(* IEC 61131-3 sources: TetherPLC/tests/compat (part 2) *)

(* ---- tc2_mc2_case.st ---- *)
PROGRAM Tc2Mc2Case
VAR
    mask   AT %QD0 : DINT;
    st     : INT;
    ax     : FB_MotionAxis;
    axH    : UDINT;
    pwr    : MC_Power;
    rst    : MC_Reset;
    sp     : MC_SetPosition;
    rpos   : MC_ReadActualPosition;
    rvel   : MC_ReadActualVelocity;
    rerr   : MC_ReadAxisError;
    rstat  : MC_ReadStatus;
    enSig  : BOOL;
    rstExec: BOOL;
    spExec : BOOL;
    spPos  : DINT;
    spMode : BOOL;
END_VAR

// Create the simulated axis once (raw FB_MotionAxis OP=1).
IF st = 0 THEN
    ax.UNITS_PER_REV := 1000;
    ax.MAX_VEL := 1000;
    ax.MAX_ACCEL := 5000;
    ax.MAX_DECEL := 5000;
    ax.POS_MIN := -100000;
    ax.POS_MAX := 100000;
    ax.HOME_OFFSET := 0;
    ax.FOLLOW_WINDOW := 3;
    ax.FLAGS := 1;
    ax.OP := 1;
    ax();
    IF ax.AXIS <> 0 AND ax.STATUS = 0 THEN
        axH := ax.AXIS;
        mask := mask + 1;
    END_IF;
    st := 1;
END_IF;

// Command/select signals derived from st (each command state is a
// single scan, giving each Execute FB exactly one rising edge).
enSig   := (st >= 1) AND (st <= 7);   // powered through the reset
rstExec := (st = 6);
spExec  := (st = 2) OR (st = 4);
spPos   := 1000;
IF st = 4 THEN spPos := 500; END_IF;
spMode  := (st = 4);

// Drive every MC wrapper each scan.
pwr(Enable := enSig, Enable_Positive := TRUE,
    Enable_Negative := TRUE, Axis := axH);
rst(Execute := rstExec, Axis := axH);
sp(Execute := spExec, Position := spPos, Mode := spMode, Axis := axH);
rpos(Enable := TRUE, Axis := axH);
rvel(Enable := TRUE, Axis := axH);
rerr(Enable := TRUE, Axis := axH);
rstat(Enable := TRUE, Axis := axH);

IF st = 1 THEN
    // MC_Power enable: wait for Status (OperationEnabled, ~2 scans)
    IF pwr.Status THEN
        mask := mask + 2;
        st := 2;
    END_IF;
ELSIF st = 2 THEN
    // absolute MC_SetPosition to 1000 fired this scan
    IF sp.Done THEN mask := mask + 4; END_IF;
    st := 3;
ELSIF st = 3 THEN
    // verify absolute position readback == 1000
    IF rpos.Valid AND rpos.Position = 1000 THEN
        mask := mask + 8;
    END_IF;
    st := 4;
ELSIF st = 4 THEN
    // relative MC_SetPosition +500 -> 1500 fired this scan
    IF sp.Done THEN mask := mask + 16; END_IF;
    st := 5;
ELSIF st = 5 THEN
    // verify relative readback == 1500 and the read FBs are valid
    IF rpos.Valid AND rpos.Position = 1500 THEN
        mask := mask + 32;
    END_IF;
    IF rvel.Valid AND rerr.Valid AND rstat.Valid THEN
        mask := mask + 64;
    END_IF;
    st := 6;
ELSIF st = 6 THEN
    // MC_Reset Execute edge -> Done (axis stays enabled)
    IF rst.Done THEN mask := mask + 128; END_IF;
    st := 7;
ELSIF st = 7 THEN
    // reset release scan; keep waiting for power to drop next
    st := 8;
ELSIF st = 8 THEN
    // enSig now FALSE: MC_Power disabled the axis; wait for
    // Status=FALSE and OperatingState=Disabled (0)
    IF NOT pwr.Status THEN
        mask := mask + 256;
        st := 9;
    END_IF;
ELSIF st = 9 THEN
    IF rstat.OperatingState = 0 THEN
        mask := mask + 512;
        st := 10;
    END_IF;
END_IF;

END_PROGRAM

(* ---- tc2_mc2_drive_case.st ---- *)
PROGRAM Tc2Mc2DriveCase
VAR
    mask   AT %QD0 : DINT;
    st     : INT;
    prevSt : INT;
    pulse  : BOOL;
    ax     : FB_MotionAxis;
    axM    : UDINT;
    axS    : UDINT;
    pwrM   : MC_Power;
    pwrS   : MC_Power;
    mvV    : MC_MoveVelocity;
    hlt    : MC_Halt;
    info   : FB_ReadDriveInfo;
    coeWr  : FB_CoEWrite;
    coeRd  : FB_CoERead;
    coeCmd : FB_CoEExecuteCommand;
    setOff : FB_SetPositionOffset;
    delOff : FB_DeletePositionOffset;
    brk    : FB_BrakeControl;
    rdPar  : FB_ReadDriveParameter;
    rdPar2 : FB_ReadDriveParameter;
    ax8kBrk : FB_CoEAX8000BrakeControl;
    ax8kTst : FB_CoEAX8000BrakeTest;
    ax8kPrk : FB_CoEAX8000ParkAxis;
    elBrk  : FB_CoEEL72xxBrakeControl;
    elSet  : FB_CoEEL72xxSetPositionOffset;
    saw    : MC_ReadFlyingSawCharacteristics;
    soeRd  : FB_SoERead;
    soeWrPw: FB_SoEWritePassword;
    soeCmd : FB_SoEExecuteCommand;
    soeCmd2: FB_SoEExecuteCommand;
    soeCmdSt: FB_SoEReadCommandState;
    soeRst : FB_SoEReset;
    ax5kV  : FB_SoEAX5000ReadActMainVoltage;
    ax5kFw : FB_SoEAX5000FirmwareUpdate;
    gv     : MC_GearInVelo;
    gp     : MC_GearInPos;
    rvelS  : MC_ReadActualVelocity;
    rposS  : MC_ReadActualPosition;
    rposM  : MC_ReadActualPosition;
    enSig  : BOOL;
    mvVEx  : BOOL;
    gvEx   : BOOL;
    gpEx   : BOOL;
    hltEx  : BOOL;
    cmdErrSeen : BOOL;
    cmdDoneSeen : BOOL;
    tog     : BOOL;
END_VAR

// Create two simulated axes (master slave0, slave slave1).
IF st = 0 THEN
    ax.UNITS_PER_REV := 1000;
    ax.MAX_VEL := 2000;
    ax.MAX_ACCEL := 8000;
    ax.MAX_DECEL := 8000;
    ax.POS_MIN := -200000;
    ax.POS_MAX := 200000;
    ax.HOME_OFFSET := 0;
    ax.FOLLOW_WINDOW := 3;
    ax.FLAGS := 1;
    ax.OP := 1; ax();
    IF ax.AXIS <> 0 THEN axM := ax.AXIS; END_IF;
    ax.OP := 1; ax();
    IF ax.AXIS <> 0 THEN axS := ax.AXIS; END_IF;
    IF axM <> 0 AND axS <> 0 THEN
        mask := mask + 1;                       // bit0: two axes
    END_IF;
    st := 1;
    prevSt := 0;
END_IF;

IF st <> prevSt THEN pulse := TRUE; ELSE pulse := FALSE; END_IF;
prevSt := st;
tog := NOT tog;   // re-pulse helper for the command-state polls

enSig  := (st >= 1) AND (st <= 29);
mvVEx  := pulse AND (st = 26);       // master velocity for gear tests
gvEx   := (st >= 27) AND (st <= 28); // velocity gear held
gpEx   := (st = 29);                 // position gear one scan
hltEx  := pulse AND (st = 30);

pwrM(Enable := enSig, Enable_Positive := TRUE, Enable_Negative := TRUE,
    Axis := axM);
pwrS(Enable := enSig, Enable_Positive := TRUE, Enable_Negative := TRUE,
    Axis := axS);
mvV(Execute := mvVEx, ContinuousUpdate := FALSE, Velocity := 400,
    Acceleration := 8000, Deceleration := 8000, Axis := axM);
hlt(Execute := hltEx, Deceleration := 8000, Axis := axM);
gv(Execute := gvEx, RatioNumerator := 2, RatioDenominator := 1,
   Acceleration := 8000, Deceleration := 8000, Master := axM, Slave := axS);
gp(Execute := gpEx, RatioNumerator := 1, RatioDenominator := 1,
   Acceleration := 8000, Deceleration := 8000, Master := axM, Slave := axS);
rvelS(Enable := TRUE, Axis := axS);
rposS(Enable := TRUE, Axis := axS);
rposM(Enable := TRUE, Axis := axM);

IF st = 1 THEN
    IF pwrM.Status AND pwrS.Status THEN
        mask := mask + 2;                       // bit1: powered
        st := 2;
    END_IF;
ELSIF st = 2 THEN
    info(Execute := pulse, Axis := axM);
    IF info.Valid AND info.State > 0 THEN
        mask := mask + 4;                       // bit2: drive info
        st := 3;
    END_IF;
ELSIF st = 3 THEN
    coeWr(Execute := pulse, Index := 16#2003, Value := 7, Axis := axM);
    IF coeWr.Done THEN
        mask := mask + 8;                       // bit3: CoE write
        st := 4;
    END_IF;
ELSIF st = 4 THEN
    coeRd(Execute := pulse, Index := 16#2003, Axis := axM);
    IF coeRd.Done AND coeRd.Value = 7 THEN
        mask := mask + 16;                      // bit4: CoE readback
        st := 5;
    END_IF;
ELSIF st = 5 THEN
    coeCmd(Execute := pulse, Command := 42, Axis := axM);
    IF coeCmd.Done THEN
        mask := mask + 32;                      // bit5: CoE command
        st := 6;
    END_IF;
ELSIF st = 6 THEN
    setOff(Execute := pulse, Position := 5000.0, Relative := FALSE,
           Feedback := 0, Memory := 0, Axis := axM);
    IF setOff.Done THEN
        mask := mask + 64;                      // bit6: pos offset
        st := 7;
    END_IF;
ELSIF st = 7 THEN
    rdPar(Execute := pulse, ParameterNumber := 16#2002, Mode := 0,
          Interval := 0, Axis := axM);
    IF rdPar.Valid AND rdPar.Value = 5000 THEN
        mask := mask + 128;                     // bit7: offset=5000
        st := 8;
    END_IF;
ELSIF st = 8 THEN
    delOff(Execute := pulse, Feedback := 0, Memory := 0, Axis := axM);
    IF delOff.Done THEN
        mask := mask + 256;                     // bit8: offset del
        st := 9;
    END_IF;
ELSIF st = 9 THEN
    brk(Execute := pulse, Mode := 3, Axis := axM);
    IF brk.Done THEN
        mask := mask + 512;                     // bit9: brake ctrl
        st := 10;
    END_IF;
ELSIF st = 10 THEN
    ax8kBrk(Execute := pulse, Mode := 1, Axis := axM);
    IF ax8kBrk.Done THEN
        mask := mask + 1024;                    // bit10: ax8k brake
        st := 11;
    END_IF;
ELSIF st = 11 THEN
    ax8kTst(Execute := pulse, Axis := axM);
    IF ax8kTst.Succeeded THEN
        mask := mask + 2048;                    // bit11: brake test
        st := 12;
    END_IF;
ELSIF st = 12 THEN
    ax8kPrk(Execute := pulse, Mode := 1, Axis := axM);
    IF ax8kPrk.Done THEN
        mask := mask + 4096;                    // bit12: ax8k park
        st := 13;
    END_IF;
ELSIF st = 13 THEN
    rdPar2(Execute := pulse, ParameterNumber := 16#2004, Mode := 0,
           Interval := 0, Axis := axM);
    IF rdPar2.Valid AND rdPar2.Value = 1 THEN
        mask := mask + 8192;                    // bit13: park=1
        st := 14;
    END_IF;
ELSIF st = 14 THEN
    elBrk(Execute := pulse, Mode := 2, Axis := axM);
    IF elBrk.Done THEN
        mask := mask + 16384;                   // bit14: el72xx brk
        st := 15;
    END_IF;
ELSIF st = 15 THEN
    elSet(Execute := pulse, Position := 7000.0, Relative := FALSE,
          Feedback := 0, Memory := 0, Axis := axM);
    IF elSet.Done THEN
        mask := mask + 32768;                   // bit15: el72xx off
        st := 16;
    END_IF;
ELSIF st = 16 THEN
    saw(Execute := pulse, Slave := axM);
    IF saw.Done AND saw.Value0 = 1000 AND saw.Value3 = 4000 THEN
        mask := mask + 65536;                   // bit16: saw charac
        st := 17;
    END_IF;
ELSIF st = 17 THEN
    soeRd(Execute := pulse, Index := 16#0135, Axis := axM);
    IF soeRd.Done AND soeRd.Value > 0.0 THEN
        mask := mask + 131072;                  // bit17: SoE status
        st := 18;
    END_IF;
ELSIF st = 18 THEN
    soeWrPw(Execute := pulse, Password := 1234, Axis := axM);
    IF soeWrPw.Done THEN
        mask := mask + 262144;                  // bit18: SoE passwd
        st := 19;
    END_IF;
ELSIF st = 19 THEN
    soeCmd(Execute := pulse, CommandId := 5, Axis := axM);
    IF soeCmd.Done THEN
        mask := mask + 524288;                  // bit19: SoE exec
        st := 20;
    END_IF;
ELSIF st = 20 THEN
    // command state polls to done (2) within the sim window;
    // tog re-pulses Execute every other scan while waiting
    IF cmdDoneSeen = FALSE THEN
        soeCmdSt(Execute := (st = 20) AND tog, Axis := axM);
        IF soeCmdSt.Done AND soeCmdSt.CommandState = 2 THEN
            cmdDoneSeen := TRUE;
            mask := mask + 1048576;             // bit20: cmd done
        END_IF;
    END_IF;
    IF cmdDoneSeen THEN st := 21; END_IF;
ELSIF st = 21 THEN
    soeCmd2(Execute := pulse, CommandId := 16#8005, Axis := axM);
    IF soeCmd2.Done THEN
        st := 22;
    END_IF;
ELSIF st = 22 THEN
    // error command (bit15) latches cmd state 3
    IF cmdErrSeen = FALSE THEN
        soeCmdSt(Execute := (st = 22) AND tog, Axis := axM);
        IF soeCmdSt.Done AND soeCmdSt.CommandState = 3 THEN
            cmdErrSeen := TRUE;
            mask := mask + 2097152;             // bit21: cmd error
        END_IF;
    END_IF;
    IF cmdErrSeen THEN st := 23; END_IF;
ELSIF st = 23 THEN
    soeRst(Execute := pulse, Axis := axM);
    IF soeRst.Done THEN
        mask := mask + 4194304;                 // bit22: SoE reset
        st := 24;
    END_IF;
ELSIF st = 24 THEN
    ax5kV(Execute := pulse, Axis := axM);
    // mains = 230 + 0.5*(sim clock steps) -> 230.0..234.5
    IF ax5kV.Done AND ax5kV.Voltage >= 230.0
       AND ax5kV.Voltage <= 234.5 THEN
        mask := mask + 8388608;                 // bit23: ax5k mains
        st := 25;
    END_IF;
ELSIF st = 25 THEN
    ax5kFw(Execute := pulse, Axis := axM);
    IF ax5kFw.Done AND ax5kFw.FirmwareRevision = 1
       AND ax5kFw.FirmwareBuild = 5 THEN
        mask := mask + 16777216;                // bit24: ax5k fw
        st := 26;
    END_IF;
ELSIF st = 26 THEN
    // master velocity move starts (mvVEx fired this scan)
    st := 27;
ELSIF st = 27 THEN
    // MC_GearInVelo 2:1: slave velocity tracks master at 2x
    IF gv.InGear AND rvelS.Valid AND
       (rvelS.Velocity >= 780) AND (rvelS.Velocity <= 820) THEN
        mask := mask + 33554432;                // bit25: gear velo
        st := 28;
    END_IF;
ELSIF st = 28 THEN
    st := 29;
ELSIF st = 29 THEN
    // MC_GearInPos 1:1: slave CSP position tracks master position
    IF gp.InGear AND rposS.Valid AND rposM.Valid AND
       (rposS.Position >= rposM.Position - 50)
       AND (rposS.Position <= rposM.Position + 50) THEN
        mask := mask + 67108864;                // bit26: gear pos
        st := 30;
    END_IF;
ELSIF st = 30 THEN
    IF NOT pwrM.Status AND NOT pwrS.Status THEN
        mask := mask + 134217728;               // bit27: powered off
        st := 31;
    END_IF;
END_IF;

END_PROGRAM

(* ---- tc2_mc2_gear_case.st ---- *)
PROGRAM Tc2Mc2GearCase
VAR
    mask   AT %QD0 : DINT;
    st     : INT;
    prevSt : INT;
    pulse  : BOOL;
    ax     : FB_MotionAxis;
    axM    : UDINT;
    axS    : UDINT;
    pwrM   : MC_Power;
    pwrS   : MC_Power;
    mvV    : MC_MoveVelocity;
    tp     : MC_TouchProbe;
    gi     : MC_GearIn;
    go     : MC_GearOut;
    hlt    : MC_Halt;
    rposM  : MC_ReadActualPosition;
    rvelM  : MC_ReadActualVelocity;
    rvelS  : MC_ReadActualVelocity;
    enSig  : BOOL;
    mvVEx  : BOOL;
    tpEx   : BOOL;
    tpTrig : BOOL;
    giEx   : BOOL;
    goEx   : BOOL;
    hltEx  : BOOL;
END_VAR

// Create the two simulated axes once (master + slave).
IF st = 0 THEN
    ax.UNITS_PER_REV := 1000;
    ax.MAX_VEL := 2000;
    ax.MAX_ACCEL := 8000;
    ax.MAX_DECEL := 8000;
    ax.POS_MIN := -200000;
    ax.POS_MAX := 200000;
    ax.HOME_OFFSET := 0;
    ax.FOLLOW_WINDOW := 3;
    ax.FLAGS := 1;
    ax.OP := 1; ax();
    IF ax.AXIS <> 0 THEN axM := ax.AXIS; END_IF;
    ax.OP := 1; ax();
    IF ax.AXIS <> 0 THEN axS := ax.AXIS; END_IF;
    IF axM <> 0 AND axS <> 0 THEN
        mask := mask + 1;                       // bit0: two axes
    END_IF;
    st := 1;
    prevSt := 0;
END_IF;

IF st <> prevSt THEN pulse := TRUE; ELSE pulse := FALSE; END_IF;
prevSt := st;

enSig  := (st >= 1) AND (st <= 7);    // both powered through st=7
mvVEx  := pulse AND (st = 2);
tpEx   := (st >= 3) AND (st <= 4);    // probe armed while moving
tpTrig := rposM.Position > 500;       // trigger as master crosses 500
giEx   := (st = 5);                   // gear held during st=5
goEx   := pulse AND (st = 6);
hltEx  := pulse AND (st = 7);

pwrM(Enable := enSig, Enable_Positive := TRUE, Enable_Negative := TRUE,
     Axis := axM);
pwrS(Enable := enSig, Enable_Positive := TRUE, Enable_Negative := TRUE,
     Axis := axS);
mvV(Execute := mvVEx, ContinuousUpdate := FALSE, Velocity := 400,
    Acceleration := 8000, Deceleration := 8000, Axis := axM);
tp(Execute := tpEx, TriggerInput := tpTrig, WindowOnly := FALSE,
   FirstPosition := 0, LastPosition := 0, Axis := axM);
gi(Execute := giEx, RatioNumerator := 2, RatioDenominator := 1,
   Acceleration := 8000, Deceleration := 8000,
   Master := axM, Slave := axS);
go(Execute := goEx, Deceleration := 8000, Slave := axS);
hlt(Execute := hltEx, Deceleration := 8000, Axis := axM);
rposM(Enable := TRUE, Axis := axM);
rvelM(Enable := TRUE, Axis := axM);
rvelS(Enable := TRUE, Axis := axS);

IF st = 1 THEN
    IF pwrM.Status AND pwrS.Status THEN
        mask := mask + 2;                       // bit1: both powered
        st := 2;
    END_IF;
ELSIF st = 2 THEN
    // master axis into velocity mode at 400
    IF mvV.InVelocity THEN
        mask := mask + 4;                       // bit2: master vel
        st := 3;
    END_IF;
ELSIF st = 3 THEN
    // MC_TouchProbe captures the position as the master crosses 500
    IF tp.Done THEN
        mask := mask + 8;                       // bit3: probe fired
        st := 4;
    END_IF;
ELSIF st = 4 THEN
    // recorded position is within one scan of the 500 trigger point
    IF tp.RecordedPosition >= 500 AND tp.RecordedPosition <= 520 THEN
        mask := mask + 16;                      // bit4: latch in window
    END_IF;
    st := 5;
ELSIF st = 5 THEN
    // MC_GearIn ratio 2/1: slave velocity tracks master at 2x = 800
    IF gi.InGear AND rvelS.Valid AND
       (rvelS.Velocity >= 780) AND (rvelS.Velocity <= 820) THEN
        mask := mask + 32;                      // bit5: geared at 800
        st := 6;
    END_IF;
ELSIF st = 6 THEN
    // gear released; MC_GearOut ramps the slave to rest
    IF go.Done THEN
        mask := mask + 64;                      // bit6: slave stopped
        st := 7;
    END_IF;
ELSIF st = 7 THEN
    // MC_Halt ramps the master to rest
    IF hlt.Done THEN
        mask := mask + 128;                     // bit7: master stopped
        st := 8;
    END_IF;
ELSIF st = 8 THEN
    // both axes powered off
    IF NOT pwrM.Status AND NOT pwrS.Status THEN
        mask := mask + 256;                     // bit8: powered off
        st := 9;
    END_IF;
END_IF;

END_PROGRAM

(* ---- tc2_mc2_modulo_case.st ---- *)
PROGRAM Tc2Mc2ModuloCase
VAR
    mask   AT %QD0 : DINT;
    st     : INT;
    prevSt : INT;
    pulse  : BOOL;
    ovrCnt : INT;
    ax     : FB_MotionAxis;
    axH    : UDINT;
    pwr    : MC_Power;
    mvMod  : MC_MoveModulo;
    mvV    : MC_MoveVelocity;
    hlt    : MC_Halt;
    ovr    : MC_SetOverride;
    rpos   : MC_ReadActualPosition;
    rvel   : MC_ReadActualVelocity;
    rstat  : MC_ReadStatus;
    rp     : MC_ReadParameter;
    rbp    : MC_ReadBoolParameter;
    wp     : MC_WriteParameter;
    wbp    : MC_WriteBoolParameter;
    enSig  : BOOL;
    mvModEx: BOOL;
    mvVEx  : BOOL;
    hltEx  : BOOL;
    wpEx   : BOOL;
    wbpEx  : BOOL;
    ovrEn  : BOOL;
    mvModP : DINT;
    mvModD : INT;
    rpNum  : UDINT;
END_VAR

// Create the simulated axis once (raw FB_MotionAxis OP=1).
IF st = 0 THEN
    ax.UNITS_PER_REV := 1000;
    ax.MAX_VEL := 2000;
    ax.MAX_ACCEL := 8000;
    ax.MAX_DECEL := 8000;
    ax.POS_MIN := -200000;
    ax.POS_MAX := 200000;
    ax.HOME_OFFSET := 0;
    ax.FOLLOW_WINDOW := 3;
    ax.FLAGS := 1;
    ax.OP := 1;
    ax();
    IF ax.AXIS <> 0 AND ax.STATUS = 0 THEN
        axH := ax.AXIS;
        mask := mask + 1;                       // bit0: axis created
    END_IF;
    st := 1;
    prevSt := 0;
END_IF;

// pulse is TRUE only on the first scan of a new phase so every
// Execute input sees exactly one rising edge per command.
IF st <> prevSt THEN pulse := TRUE; ELSE pulse := FALSE; END_IF;
prevSt := st;

enSig   := (st >= 1) AND (st <= 11);  // powered through the commands
mvModEx := pulse AND ((st = 2) OR (st = 4));
mvModP  := 270; IF st = 4 THEN mvModP := 90; END_IF;
mvModD  := 0;   IF st = 4 THEN mvModD := 1; END_IF;
mvVEx   := pulse AND (st = 9);
hltEx   := pulse AND (st = 11);
wpEx    := pulse AND (st = 6);
wbpEx   := pulse AND (st = 8);
ovrEn   := (st = 10);
rpNum   := 16#6065; IF st = 8 THEN rpNum := 16#607C; END_IF;

// Drive every MC wrapper each scan. ovr is called before hlt so a
// simultaneous override-restore does not clobber the halt target.
pwr(Enable := enSig, Enable_Positive := TRUE,
    Enable_Negative := TRUE, Axis := axH);
mvMod(Execute := mvModEx, Position := mvModP, Velocity := 2000,
      Acceleration := 8000, Deceleration := 8000, Direction := mvModD,
      ModuloFactor := 360, Axis := axH);
mvV(Execute := mvVEx, ContinuousUpdate := FALSE, Velocity := 400,
    Acceleration := 8000, Deceleration := 8000, Axis := axH);
ovr(Enable := ovrEn, VelFactor := 50, Axis := axH);
hlt(Execute := hltEx, Deceleration := 8000, Axis := axH);
wp(Execute := wpEx, ParameterNumber := 16#6065, Value := 30, Axis := axH);
wbp(Execute := wbpEx, ParameterNumber := 16#607C, Value := TRUE, Axis := axH);
rp(Enable := TRUE, ParameterNumber := rpNum, Axis := axH);
rbp(Enable := TRUE, ParameterNumber := 16#6041, Axis := axH);
rpos(Enable := TRUE, Axis := axH);
rvel(Enable := TRUE, Axis := axH);
rstat(Enable := TRUE, Axis := axH);

IF st = 1 THEN
    IF pwr.Status THEN
        mask := mask + 2;                       // bit1: powered
        st := 2;
    END_IF;
ELSIF st = 2 THEN
    // MC_MoveModulo shortest to 270deg from 0 -> lands at -90
    IF mvMod.Done THEN
        mask := mask + 4;                       // bit2: modulo done
        st := 3;
    END_IF;
ELSIF st = 3 THEN
    IF rpos.Valid AND (rpos.Position >= -93) AND (rpos.Position <= -87) THEN
        mask := mask + 8;                       // bit3: pos==-90
    END_IF;
    st := 4;
ELSIF st = 4 THEN
    // MC_MoveModulo positive-direction to 90deg from -90 -> lands 90
    IF mvMod.Done THEN
        mask := mask + 16;                      // bit4: modulo done
        st := 5;
    END_IF;
ELSIF st = 5 THEN
    IF rpos.Valid AND (rpos.Position >= 87) AND (rpos.Position <= 93) THEN
        mask := mask + 32;                      // bit5: pos==90
    END_IF;
    st := 6;
ELSIF st = 6 THEN
    // MC_WriteParameter: following window 0x6065 := 30
    IF wp.Done THEN
        mask := mask + 64;                      // bit6: write done
        st := 7;
    END_IF;
ELSIF st = 7 THEN
    // MC_ReadParameter(0x6065)==30 and MC_ReadBoolParameter(0x6041)
    IF rp.Valid AND rp.Value = 30 AND rbp.Valid AND rbp.Value THEN
        mask := mask + 128;                     // bit7: param readback
        st := 8;
    END_IF;
ELSIF st = 8 THEN
    // MC_WriteBoolParameter: home offset 0x607C := 1, read back ==1
    IF wbp.Done AND rp.Valid AND rp.Value = 1 THEN
        mask := mask + 256;                     // bit8: bool param rt
        st := 9;
    END_IF;
ELSIF st = 9 THEN
    // MC_MoveVelocity ramps to 400 and holds
    IF mvV.InVelocity THEN
        st := 10;
        ovrCnt := 0;
    END_IF;
ELSIF st = 10 THEN
    // MC_SetOverride 50% halves the velocity target to ~200; the
    // axis should report ContinuousMotion (PLCopen state 4)
    ovrCnt := ovrCnt + 1;
    IF ovrCnt > 40 THEN
        IF rvel.Valid AND (rvel.Velocity >= 190) AND (rvel.Velocity <= 210)
           AND rstat.OperatingState = 4 THEN
            mask := mask + 512;                 // bit9: override+state
        END_IF;
        st := 11;
    END_IF;
ELSIF st = 11 THEN
    // override releases, MC_Halt ramps to rest and stays enabled
    IF hlt.Done AND rstat.OperatingState = 1 THEN
        mask := mask + 1024;                    // bit10: halt+standstill
        st := 12;
    END_IF;
ELSIF st = 12 THEN
    // MC_Power disable: wait for Status to drop
    IF NOT pwr.Status THEN
        mask := mask + 2048;                    // bit11: powered off
        st := 13;
    END_IF;
END_IF;

END_PROGRAM

(* ---- tc2_mc2_motion_case.st ---- *)
PROGRAM Tc2Mc2MotionCase
VAR
    mask   AT %QD0 : DINT;
    st     : INT;
    prevSt : INT;
    pulse  : BOOL;
    jogCnt : INT;
    ax     : FB_MotionAxis;
    axH    : UDINT;
    pwr    : MC_Power;
    mvA    : MC_MoveAbsolute;
    mvR    : MC_MoveRelative;
    mvV    : MC_MoveVelocity;
    stp    : MC_Stop;
    hlt    : MC_Halt;
    hom    : MC_Home;
    jog    : MC_Jog;
    rpos   : MC_ReadActualPosition;
    enSig  : BOOL;
    mvAEx  : BOOL;
    mvREx  : BOOL;
    mvVEx  : BOOL;
    stpEx  : BOOL;
    hltEx  : BOOL;
    homEx  : BOOL;
    jogF   : BOOL;
END_VAR

// Create the simulated axis once (raw FB_MotionAxis OP=1).
IF st = 0 THEN
    ax.UNITS_PER_REV := 1000;
    ax.MAX_VEL := 2000;
    ax.MAX_ACCEL := 8000;
    ax.MAX_DECEL := 8000;
    ax.POS_MIN := -200000;
    ax.POS_MAX := 200000;
    ax.HOME_OFFSET := 0;
    ax.FOLLOW_WINDOW := 3;
    ax.FLAGS := 1;
    ax.OP := 1;
    ax();
    IF ax.AXIS <> 0 AND ax.STATUS = 0 THEN
        axH := ax.AXIS;
        mask := mask + 1;                       // bit0: axis created
    END_IF;
    st := 1;
    prevSt := 0;
END_IF;

// pulse is TRUE only on the first scan of a new phase so every
// Execute input sees exactly one rising edge per command.
IF st <> prevSt THEN pulse := TRUE; ELSE pulse := FALSE; END_IF;
prevSt := st;

// Level/edge inputs derived from the current phase.
enSig := (st >= 1) AND (st <= 11);   // powered through the commands
mvAEx := pulse AND (st = 2);
mvREx := pulse AND (st = 4);
mvVEx := pulse AND ((st = 6) OR (st = 8));
stpEx := pulse AND (st = 7);
hltEx := pulse AND (st = 9);
homEx := pulse AND (st = 10);
jogF  := (st = 11) AND (jogCnt < 60);

// Drive every MC wrapper each scan.
pwr(Enable := enSig, Enable_Positive := TRUE,
    Enable_Negative := TRUE, Axis := axH);
mvA(Execute := mvAEx, Position := 1000, Velocity := 2000,
    Acceleration := 8000, Deceleration := 8000, Axis := axH);
mvR(Execute := mvREx, Distance := 500, Velocity := 2000,
    Acceleration := 8000, Deceleration := 8000, Axis := axH);
mvV(Execute := mvVEx, ContinuousUpdate := FALSE, Velocity := 400,
    Acceleration := 8000, Deceleration := 8000, Axis := axH);
stp(Execute := stpEx, Deceleration := 8000, Axis := axH);
hlt(Execute := hltEx, Deceleration := 8000, Axis := axH);
hom(Execute := homEx, Position := 0, Velocity := 2000,
    Acceleration := 8000, Deceleration := 8000, Axis := axH);
jog(JogForward := jogF, JogBackwards := FALSE, Velocity := 400,
    Axis := axH);
rpos(Enable := TRUE, Axis := axH);

IF st = 1 THEN
    // MC_Power enable: wait for Status (OperationEnabled)
    IF pwr.Status THEN
        mask := mask + 2;                       // bit1: powered
        st := 2;
    END_IF;
ELSIF st = 2 THEN
    // MC_MoveAbsolute to 1000
    IF mvA.Done THEN
        mask := mask + 4;                       // bit2: abs move done
        st := 3;
    END_IF;
ELSIF st = 3 THEN
    // verify absolute position near 1000 (within follow window)
    IF rpos.Valid AND (rpos.Position >= 997) AND (rpos.Position <= 1003) THEN
        mask := mask + 8;                       // bit3: pos==1000
    END_IF;
    st := 4;
ELSIF st = 4 THEN
    // MC_MoveRelative +500 -> ~1500
    IF mvR.Done THEN
        mask := mask + 16;                      // bit4: rel move done
        st := 5;
    END_IF;
ELSIF st = 5 THEN
    IF rpos.Valid AND (rpos.Position >= 1497) AND (rpos.Position <= 1503) THEN
        mask := mask + 32;                      // bit5: pos==1500
    END_IF;
    st := 6;
ELSIF st = 6 THEN
    // MC_MoveVelocity ramps to 400 and holds
    IF mvV.InVelocity THEN
        mask := mask + 64;                      // bit6: in velocity
        st := 7;
    END_IF;
ELSIF st = 7 THEN
    // MC_Stop quick-stop locks the axis at rest
    IF stp.Done THEN
        mask := mask + 128;                     // bit7: stopped
        st := 8;
    END_IF;
ELSIF st = 8 THEN
    // re-issue MC_MoveVelocity (recovers from quick stop)
    IF mvV.InVelocity THEN
        st := 9;
    END_IF;
ELSIF st = 9 THEN
    // MC_Halt ramps to rest but keeps the axis enabled
    IF hlt.Done THEN
        mask := mask + 256;                     // bit8: halted
        st := 10;
    END_IF;
ELSIF st = 10 THEN
    // MC_Home moves back to the home offset (0)
    IF hom.Done THEN
        mask := mask + 512;                     // bit9: homed
        st := 11;
        jogCnt := 0;
    END_IF;
ELSIF st = 11 THEN
    // MC_Jog forward ~60 scans then release; Done on rest
    jogCnt := jogCnt + 1;
    IF jog.Done AND rpos.Valid AND (rpos.Position > 50) THEN
        mask := mask + 1024;                    // bit10: jog done
        mask := mask + 2048;                    // bit11: jogged +pos
        st := 12;
    END_IF;
ELSIF st = 12 THEN
    // MC_Power disable: wait for Status to drop
    IF NOT pwr.Status THEN
        mask := mask + 4096;                    // bit12: powered off
        st := 13;
    END_IF;
END_IF;

END_PROGRAM

(* ---- tc2_mc2_probe_case.st ---- *)
PROGRAM Tc2Mc2ProbeCase
VAR
    mask   AT %QD0 : DINT;
    st     : INT;
    prevSt : INT;
    pulse  : BOOL;
    ax     : FB_MotionAxis;
    axM    : UDINT;
    pwr    : MC_Power;
    sp     : MC_SetPosition;
    tp     : MC_TouchProbe;
    ab     : MC_AbortTrigger;
    rpos   : MC_ReadActualPosition;
    enSig  : BOOL;
    spEx   : BOOL;
    tpEx   : BOOL;
    abEx   : BOOL;
    tpTrig : BOOL;
    abSeen : BOOL;
    abDoneSeen : BOOL;
    disarmed   : BOOL;
END_VAR

// Create one simulated axis.
IF st = 0 THEN
    ax.UNITS_PER_REV := 1000;
    ax.MAX_VEL := 2000;
    ax.MAX_ACCEL := 8000;
    ax.MAX_DECEL := 8000;
    ax.POS_MIN := -200000;
    ax.POS_MAX := 200000;
    ax.HOME_OFFSET := 0;
    ax.FOLLOW_WINDOW := 3;
    ax.FLAGS := 1;
    ax.OP := 1; ax();
    IF ax.AXIS <> 0 THEN axM := ax.AXIS; END_IF;
    IF axM <> 0 THEN
        mask := mask + 1;                       // bit0: axis created
    END_IF;
    st := 1;
    prevSt := 0;
END_IF;

IF st <> prevSt THEN pulse := TRUE; ELSE pulse := FALSE; END_IF;
prevSt := st;

enSig  := (st >= 1) AND (st <= 10);   // powered through st=10
spEx   := pulse AND (st = 2);        // preset position 1000
tpEx   := pulse AND (st = 5 OR st = 9);  // arm, later re-arm
abEx   := pulse AND (st = 7);        // abort the armed probe
tpTrig := (st >= 9);                 // trigger edge on re-arm scan

pwr(Enable := enSig, Enable_Positive := TRUE, Enable_Negative := TRUE,
    Axis := axM);
sp(Execute := spEx, Position := 1000, Mode := FALSE, Axis := axM);
tp(Execute := tpEx, TriggerInput := tpTrig, WindowOnly := FALSE,
   FirstPosition := 0, LastPosition := 0, Axis := axM);
ab(Execute := abEx, TriggerInput := FALSE, Axis := axM);
rpos(Enable := TRUE, Axis := axM);

IF st = 1 THEN
    IF pwr.Status THEN
        mask := mask + 2;                       // bit1: powered
        st := 2;
    END_IF;
ELSIF st = 2 THEN
    // MC_SetPosition edge writes 1000; Done pulses on this scan
    IF sp.Done THEN
        mask := mask + 256;                     // bit8: pos preset
        st := 3;
    END_IF;
ELSIF st = 3 THEN
    st := 4;
ELSIF st = 4 THEN
    st := 5;
ELSIF st = 5 THEN
    // probe armed this scan (Execute edge)
    st := 6;
ELSIF st = 6 THEN
    IF tp.Busy THEN
        mask := mask + 4;                       // bit2: probe armed
        st := 7;
    END_IF;
ELSIF st = 7 THEN
    // MC_AbortTrigger Execute edge writes the abort request
    st := 8;
ELSIF st = 8 THEN
    // wait until the armed probe consumes the abort (may take an
    // extra scan over Tether IO)
    IF tp.CommandAborted AND NOT abSeen THEN
        abSeen := TRUE;
        mask := mask + 8;                       // bit3: probe aborted
    END_IF;
    IF ab.Done AND NOT abDoneSeen THEN
        abDoneSeen := TRUE;
        mask := mask + 16;                      // bit4: abort Done
    END_IF;
    IF NOT tp.Busy AND NOT disarmed THEN
        disarmed := TRUE;
        mask := mask + 32;                      // bit5: probe idle
    END_IF;
    IF abSeen AND abDoneSeen AND disarmed THEN
        st := 9;
    END_IF;
ELSIF st = 9 THEN
    // re-arm + trigger edge in the same scan: probe captures pos
    IF tp.Done THEN
        mask := mask + 64;                      // bit6: captured
        st := 10;
    END_IF;
ELSIF st = 10 THEN
    // recorded position equals the preset axis position
    IF rpos.Valid AND tp.RecordedPosition = rpos.Position
       AND tp.RecordedPosition = 1000 THEN
        mask := mask + 128;                     // bit7: pos matches
    END_IF;
    st := 11;
ELSIF st = 11 THEN
    // power off
    IF NOT pwr.Status THEN
        mask := mask + 512;                     // bit9: powered off
        st := 12;
    END_IF;
END_IF;

END_PROGRAM

(* ---- tc2_mc2_xfc_case.st ---- *)
// e2e for compat/tc2/tc2_mc2_xfc.st — XFC kinematics, cams,
// digital cam switches and touch probe over a simulated axis.
// Mask bits (expected 0xFFFF):
//  0 axis created   1 powered        2 pos preset     3 vel reached
//  4 posAtTime#1    5 posAtTime#2    6 timeOfPos      7 timeToPos
//  8 timeToModulo   9 extendDcTime  10 curDcTime     11 camPos early-off
// 12 cams crossed  13 timeCam fired+cleared
// 14 breakcam+dcs state  15 touchprobe done+position
PROGRAM Tc2Mc2XfcCase
VAR
    mask   AT %QD0 : DINT;
    st     : INT;
    prevSt : INT;
    pulse  : BOOL;

    ax     : FB_MotionAxis;
    rd     : FB_MotionAxis;
    axM    : UDINT;

    pwr    : MC_Power;
    sp     : MC_SetPosition;
    mv     : MC_MoveVelocity;
    stp    : MC_Stop;

    curTm  : XFC_GetCurDcTaskTime;
    posAt  : XFC_PositionAtTime;
    posAtB : XFC_PositionAtTime;
    timOf  : XFC_TimeOfPosition;
    timTo  : XFC_TimeToPosition;
    timMod : XFC_TimeToModuloPosition;
    timMod2: XFC_TimeToModuloPosition;
    extDc  : XFC_ExtendDcTime;
    camPos : XFC_PositionCam;
    camTim : XFC_TimeCam;
    camBrk : XFC_BreakCam;
    dcs    : MC_DigitalCamSwitch;
    dcsMe  : MC_DigitalCamSwitch_MultiEdge;
    prb    : XFC_TouchProbe;

    enSig  : BOOL;
    mvEx   : BOOL;
    spEx   : BOOL;
    stpEx  : BOOL;
    prbEx  : BOOL;
    prbTrig: BOOL;

    posL   : LREAL;
    velL   : LREAL;
    basePos: LREAL;
    camOn  : LREAL;
    camOff : LREAL;
    t0     : UDINT;
    dDt    : DINT;
    exp    : LREAL;
    posAtDcA : UDINT;
    posAtDcB : UDINT;
    timOfPos : LREAL;
    timToPos : LREAL;
    timModPos  : LREAL;
    timModPos2 : LREAL;

    camOnSeen  : BOOL;
    dcsOnSeen  : BOOL;
    dcsMeOnSeen: BOOL;
    tcamOn     : BOOL;
    prbDone    : BOOL;
    prbRec     : LREAL;
END_VAR

// ---- per-scan FB calls ----------------------------------------------
IF st <> prevSt THEN pulse := TRUE; ELSE pulse := FALSE; END_IF;
prevSt := st;

IF axM <> 0 THEN
    rd.AXIS := axM; rd.OP := 6; rd();
END_IF;
posL := DINT_TO_LREAL(rd.POS_ACTUAL);
velL := DINT_TO_LREAL(rd.VEL_ACTUAL);

curTm();
// kinematic FBs run every scan so their internal clocks share the
// program-start epoch; query inputs are preset one stage ahead
posAt(DcTime := posAtDcA, Axis := axM);
posAtB(DcTime := posAtDcB, Axis := axM);
timOf(Position := timOfPos, Axis := axM);
timTo(Position := timToPos, Axis := axM);
timMod(Position := timModPos, ModuloFactor := 4000.0, Axis := axM);
timMod2(Position := timModPos2, ModuloFactor := 4000.0, Axis := axM);

camPos(FirstOnPosition := camOn, LastOnPosition := camOff,
       Modulo := FALSE, ModuloFactor := 0.0, Axis := axM);
camTim(FirstOnPosition := camOn + 100.0, Duration := 0.02,
       Modulo := FALSE, ModuloFactor := 0.0, Axis := axM);
camBrk(BreakRelease := TRUE, Axis := axM);
dcs(Enable := TRUE, FirstOnPosition := camOn, LastOnPosition := camOff,
    Modulo := FALSE, ModuloFactor := 0.0, Axis := axM);
dcsMe(Enable := TRUE, FirstOnPosition := camOn, LastOnPosition := camOff,
      Modulo := FALSE, ModuloFactor := 0.0, Axis := axM);

IF camPos.Output THEN camOnSeen := TRUE; END_IF;
IF dcs.Output THEN dcsOnSeen := TRUE; END_IF;
IF dcsMe.Output THEN dcsMeOnSeen := TRUE; END_IF;
IF camTim.Output THEN tcamOn := TRUE; END_IF;
IF prb.Done THEN
    prbDone := TRUE;
    prbRec := prb.RecordedPosition;
END_IF;

// ---- stage inputs ----------------------------------------------------
enSig   := (st >= 1) AND (st <= 30);
mvEx    := pulse AND (st = 5);
spEx    := pulse AND (st = 2);
stpEx   := pulse AND (st = 12);
prbEx   := (st >= 15);
prbTrig := (st >= 17);

pwr(Enable := enSig, Enable_Positive := TRUE, Enable_Negative := TRUE,
    Axis := axM);
sp(Execute := spEx, Position := 0, Mode := FALSE, Axis := axM);
mv(Execute := mvEx, ContinuousUpdate := FALSE, Velocity := 5000,
   Acceleration := 50000, Deceleration := 50000, Axis := axM);
stp(Execute := stpEx, Deceleration := 50000, Axis := axM);
prb(Execute := prbEx, TriggerInput := prbTrig, Axis := axM);

// ---- stages ----------------------------------------------------------
IF st = 0 THEN
    ax.UNITS_PER_REV := 1000;
    ax.MAX_VEL := 10000;
    ax.MAX_ACCEL := 50000;
    ax.MAX_DECEL := 50000;
    ax.POS_MIN := -2000000;
    ax.POS_MAX := 2000000;
    ax.HOME_OFFSET := 0;
    ax.FOLLOW_WINDOW := 3;
    ax.FLAGS := 1;
    ax.OP := 1; ax();
    IF ax.AXIS <> 0 THEN axM := ax.AXIS; END_IF;
    IF axM <> 0 THEN
        mask := mask + 1;                       // bit0
    END_IF;
    st := 1;
ELSIF st = 1 THEN
    IF pwr.Status THEN
        mask := mask + 2;                       // bit1
        st := 2;
    END_IF;
ELSIF st = 2 THEN
    IF sp.Done THEN
        mask := mask + 4;                       // bit2
        st := 3;
    END_IF;
ELSIF st = 3 THEN
    st := 4;
ELSIF st = 4 THEN
    st := 5;
ELSIF st = 5 THEN
    st := 6;
ELSIF st = 6 THEN
    // wait for the velocity ramp (>2500 of 5000 u/s)
    IF rd.VEL_ACTUAL > 2500 THEN
        mask := mask + 8;                       // bit3
        st := 7;
    END_IF;
ELSIF st = 7 THEN
    basePos := posL;
    camOn := basePos + 200.0;
    camOff := basePos + 500.0;
    t0 := curTm.DcTime;
    posAtDcA := t0;
    posAtDcB := t0 + 300000000;
    timOfPos := posL + 500.0;
    timToPos := posL + 500.0;
    timModPos := posL + 500.0;
    timModPos2 := posL - 3500.0;
    st := 8;
ELSIF st = 8 THEN
    // kinematic FB outputs from the per-scan calls (inputs preset
    // at st7 against the shared clock epoch)
    dDt := UDINT_TO_DINT(posAtDcA - curTm.DcTime);
    exp := posL + velL * DINT_TO_LREAL(dDt) / 1000000000.0;
    IF posAt.Error = FALSE AND
       (posAt.Position - exp > -150.0) AND
       (posAt.Position - exp < 150.0) THEN
        mask := mask + 16;                      // bit4
    END_IF;
    dDt := UDINT_TO_DINT(posAtDcB - curTm.DcTime);
    exp := posL + velL * DINT_TO_LREAL(dDt) / 1000000000.0;
    IF posAtB.Error = FALSE AND
       (posAtB.Position - exp > -150.0) AND
       (posAtB.Position - exp < 150.0) THEN
        mask := mask + 32;                      // bit5
    END_IF;
    // time-of / time-to position: +500 u at ~5000 u/s ~ 1e8 ns
    dDt := UDINT_TO_DINT(timOf.DcTime - t0);
    IF timOf.Error = FALSE AND dDt > 30000000 AND dDt < 300000000 THEN
        mask := mask + 64;                      // bit6
    END_IF;
    IF timTo.Error = FALSE AND timTo.Duration > 30000000
       AND timTo.Duration < 300000000 THEN
        mask := mask + 128;                     // bit7
    END_IF;
    IF timMod.Error = FALSE AND timMod2.Error = FALSE
       AND timMod.Duration > 30000000 AND timMod.Duration < 300000000
       AND timMod2.Duration > 30000000 AND timMod2.Duration < 300000000 THEN
        mask := mask + 256;                     // bit8
    END_IF;
    extDc(DcTime32 := 501234, RefDcTime := 500000);
    IF extDc.DeltaNs = 1234 THEN
        mask := mask + 512;                     // bit9
    END_IF;
    IF curTm.DcTime <> 0 THEN
        mask := mask + 1024;                    // bit10
    END_IF;
    IF NOT camPos.Output THEN
        mask := mask + 2048;                     // bit11: cam still off
    END_IF;
    st := 9;
ELSIF st = 9 THEN
    st := 10;
ELSIF st = 10 THEN
    st := 11;
ELSIF st = 11 THEN
    // move still running; cam windows are crossed here
    st := 12;
ELSIF st = 12 THEN
    st := 13;
ELSIF st = 13 THEN
    // wait for the stop to complete
    IF rd.VEL_ACTUAL < 50 THEN
        st := 14;
    END_IF;
ELSIF st = 14 THEN
    st := 15;
ELSIF st = 15 THEN
    st := 16;
ELSIF st = 16 THEN
    st := 17;
ELSIF st = 17 THEN
    IF camOnSeen AND dcsOnSeen AND dcsMeOnSeen THEN
        mask := mask + 4096;                     // bit12
    END_IF;
    IF tcamOn AND NOT camTim.Output THEN
        mask := mask + 8192;                     // bit13
    END_IF;
    IF camBrk.Output AND dcs.InOperation
       AND dcsMe.InOperation THEN
        mask := mask + 16384;                    // bit14
    END_IF;
    st := 18;
ELSIF st = 18 THEN
    st := 19;
ELSIF st = 19 THEN
    IF prbDone AND (prbRec - posL > -200.0)
       AND (prbRec - posL < 200.0) THEN
        mask := mask + 32768;                    // bit15
    END_IF;
    st := 20;
ELSIF st = 20 THEN
    st := 21;
END_IF;

END_PROGRAM

(* ---- tc2_modbusrtu_case.st ---- *)
PROGRAM Tc2ModbusRtuCase
VAR
    mask      AT %QD0   : DINT;
    st        : INT;
    scan_n    : UDINT;
    rregs     : FB_MBRtuReadRegs;
    wsreg     : FB_MBRtuWriteSingleReg;
    wregs     : FB_MBRtuWriteRegs;
    rcoils    : FB_MBRtuReadCoils;
    rbad      : FB_MBRtuReadRegs;
    rwregs    : FB_MBRtuReadWriteRegs;
    wsrc      : ARRAY[0..255] OF BYTE;
END_VAR

// autonomous Modbus RTU sequence against tests/compat/
// modbus_rtu_test_server.py over a pty pair: read regs ->
// write single reg -> write regs -> read coils -> exception
// read -> read/write regs. sDevice is substituted by the test
// script with the pty slave path.
wsrc[0] := 16#12;
wsrc[1] := 16#34;

rregs(bExecute := st = 0, tTimeout := T#5s,
      sDevice := '__PTY_SLAVE__', nBaud := 9600,
      nParity := 0, nDataBits := 8, nStopBits := 1,
      nUnitID := 1, nQuantity := 2, nMBAddr := 0,
      cbLength := 256);
wsreg(bExecute := st = 1, tTimeout := T#5s,
      sDevice := '__PTY_SLAVE__', nBaud := 9600,
      nParity := 0, nDataBits := 8, nStopBits := 1,
      nUnitID := 1, nMBAddr := 0, nValue := 16#BEEF);
wregs(bExecute := st = 2, tTimeout := T#5s,
      sDevice := '__PTY_SLAVE__', nBaud := 9600,
      nParity := 0, nDataBits := 8, nStopBits := 1,
      nUnitID := 1, nQuantity := 2, nMBAddr := 0,
      cbLength := 4, pSrcData := wsrc);
rcoils(bExecute := st = 3, tTimeout := T#5s,
       sDevice := '__PTY_SLAVE__', nBaud := 9600,
       nParity := 0, nDataBits := 8, nStopBits := 1,
       nUnitID := 1, nQuantity := 8, nMBAddr := 0,
       cbLength := 256);
rbad(bExecute := st = 4, tTimeout := T#5s,
     sDevice := '__PTY_SLAVE__', nBaud := 9600,
     nParity := 0, nDataBits := 8, nStopBits := 1,
     nUnitID := 1, nQuantity := 2, nMBAddr := 99,
     cbLength := 256);
rwregs(bExecute := st = 5, tTimeout := T#5s,
       sDevice := '__PTY_SLAVE__', nBaud := 9600,
       nParity := 0, nDataBits := 8, nStopBits := 1,
       nUnitID := 1, nReadQuantity := 2, nMBReadAddr := 0,
       nWriteQuantity := 1, nMBWriteAddr := 0,
       cbDestLength := 256, cbSrcLength := 2,
       pSrcData := wsrc);

IF st = 0 AND rregs.bDone THEN
    // func3 resp PDU data = bytecount + reg bytes
    IF rregs.bError = FALSE AND rregs.cbRead = 5 AND
       rregs.pData[0] = 4 AND rregs.pData[1] = 16#10 AND
       rregs.pData[2] = 16#00 AND rregs.pData[3] = 16#10 AND
       rregs.pData[4] = 16#01 THEN
        mask := mask + 1;
    END_IF;
    st := 1;
ELSIF st = 1 AND wsreg.bDone THEN
    IF wsreg.bError = FALSE AND wsreg.nErrId = 0 THEN
        mask := mask + 2;
    END_IF;
    st := 2;
ELSIF st = 2 AND wregs.bDone THEN
    IF wregs.bError = FALSE AND wregs.nErrId = 0 THEN
        mask := mask + 4;
    END_IF;
    st := 3;
ELSIF st = 3 AND rcoils.bDone THEN
    // func1 resp = bytecount(1) + 0xA5
    IF rcoils.bError = FALSE AND rcoils.cbRead = 2 AND
       rcoils.pData[0] = 1 AND rcoils.pData[1] = 16#A5 THEN
        mask := mask + 8;
    END_IF;
    st := 4;
ELSIF st = 4 AND rbad.bDone THEN
    // addr 99 -> server exception 2 -> nErrId = 16#8002
    IF rbad.bError = TRUE AND rbad.nErrId = 16#8002 THEN
        mask := mask + 16;
    END_IF;
    st := 5;
ELSIF st = 5 AND rwregs.bDone THEN
    IF rwregs.bError = FALSE AND rwregs.cbRead = 5 AND
       rwregs.pDestData[0] = 4 AND rwregs.pDestData[1] = 16#10 AND
       rwregs.pDestData[4] = 16#01 THEN
        mask := mask + 32;
    END_IF;
    st := 6;
END_IF;

scan_n := scan_n + 1;
END_PROGRAM

(* ---- tc2_modbussrv_case.st ---- *)
PROGRAM Tc2ModbusSrvCase
VAR
    mask      AT %QD0   : DINT;
    st        : INT;
    scan_n    : UDINT;
    rregs     : FB_MBReadRegs;
    wsreg     : FB_MBWriteSingleReg;
    wregs     : FB_MBWriteRegs;
    rcoils    : FB_MBReadCoils;
    rbad      : FB_MBReadRegs;
    rwregs    : FB_MBReadWriteRegs;
    wsrc      : ARRAY[0..255] OF BYTE;
END_VAR

// autonomous Modbus TCP sequence against tests/compat/
// modbus_test_server.py: read regs -> write single reg ->
// write regs -> read coils -> exception read -> read/write regs.
// Each state's bExecute is high only while st equals its index,
// giving every FB one rising edge.
wsrc[0] := 16#12;
wsrc[1] := 16#34;

rregs(bExecute := st = 0, tTimeout := T#5s,
      sHost := '127.0.0.1', nTCPPort := 15088,
      nUnitID := 16#FF, nQuantity := 2, nMBAddr := 0,
      cbLength := 256);
wsreg(bExecute := st = 1, tTimeout := T#5s,
      sHost := '127.0.0.1', nTCPPort := 15088,
      nUnitID := 16#FF, nMBAddr := 0, nValue := 16#BEEF);
wregs(bExecute := st = 2, tTimeout := T#5s,
      sHost := '127.0.0.1', nTCPPort := 15088,
      nUnitID := 16#FF, nQuantity := 2, nMBAddr := 0,
      cbLength := 4, pSrcData := wsrc);
rcoils(bExecute := st = 3, tTimeout := T#5s,
       sHost := '127.0.0.1', nTCPPort := 15088,
       nUnitID := 16#FF, nQuantity := 8, nMBAddr := 0,
       cbLength := 256);
rbad(bExecute := st = 4, tTimeout := T#5s,
     sHost := '127.0.0.1', nTCPPort := 15088,
     nUnitID := 16#FF, nQuantity := 2, nMBAddr := 99,
     cbLength := 256);
rwregs(bExecute := st = 5, tTimeout := T#5s,
       sHost := '127.0.0.1', nTCPPort := 15088,
       nUnitID := 16#FF, nReadQuantity := 2, nMBReadAddr := 0,
       nWriteQuantity := 1, nMBWriteAddr := 0,
       cbDestLength := 256, cbSrcLength := 2,
       pSrcData := wsrc);

IF st = 0 AND rregs.bDone THEN
    // func3 resp PDU data = bytecount + reg bytes
    IF rregs.bError = FALSE AND rregs.cbRead = 5 AND
       rregs.pData[0] = 4 AND rregs.pData[1] = 16#10 AND
       rregs.pData[2] = 16#00 AND rregs.pData[3] = 16#10 AND
       rregs.pData[4] = 16#01 THEN
        mask := mask + 1;
    END_IF;
    st := 1;
ELSIF st = 1 AND wsreg.bDone THEN
    IF wsreg.bError = FALSE AND wsreg.nErrId = 0 THEN
        mask := mask + 2;
    END_IF;
    st := 2;
ELSIF st = 2 AND wregs.bDone THEN
    IF wregs.bError = FALSE AND wregs.nErrId = 0 THEN
        mask := mask + 4;
    END_IF;
    st := 3;
ELSIF st = 3 AND rcoils.bDone THEN
    // func1 resp = bytecount(1) + 0xA5
    IF rcoils.bError = FALSE AND rcoils.cbRead = 2 AND
       rcoils.pData[0] = 1 AND rcoils.pData[1] = 16#A5 THEN
        mask := mask + 8;
    END_IF;
    st := 4;
ELSIF st = 4 AND rbad.bDone THEN
    // addr 99 -> server exception 2 -> nErrId = 16#8002
    IF rbad.bError = TRUE AND rbad.nErrId = 16#8002 THEN
        mask := mask + 16;
    END_IF;
    st := 5;
ELSIF st = 5 AND rwregs.bDone THEN
    IF rwregs.bError = FALSE AND rwregs.cbRead = 5 AND
       rwregs.pDestData[0] = 4 AND rwregs.pDestData[1] = 16#10 AND
       rwregs.pDestData[4] = 16#01 THEN
        mask := mask + 32;
    END_IF;
    st := 6;
END_IF;

scan_n := scan_n + 1;
END_PROGRAM

(* ---- tc2_modbussrv_udp_case.st ---- *)
PROGRAM Tc2ModbusSrvUdpCase
VAR
    mask      AT %QD0   : DINT;
    st        : INT;
    scan_n    : UDINT;
    rregs     : FB_MBUdpReadRegs;
    wsreg     : FB_MBUdpWriteSingleReg;
    rcoils    : FB_MBUdpReadCoils;
    rbad      : FB_MBUdpReadRegs;
    rwregs    : FB_MBUdpReadWriteRegs;
    wsrc      : ARRAY[0..255] OF BYTE;
END_VAR

// autonomous Modbus UDP sequence against tests/compat/
// modbus_test_server.py (UDP peer on port 15089): read regs ->
// write single reg -> read coils -> exception read -> read/write
// regs. Each state's bExecute is high only while st equals its
// index, giving every FB one rising edge.
wsrc[0] := 16#12;
wsrc[1] := 16#34;

rregs(bExecute := st = 0, tTimeout := T#5s,
      sHost := '127.0.0.1', nTCPPort := 15089,
      nUnitID := 16#FF, nQuantity := 2, nMBAddr := 0,
      cbLength := 256);
wsreg(bExecute := st = 1, tTimeout := T#5s,
      sHost := '127.0.0.1', nTCPPort := 15089,
      nUnitID := 16#FF, nMBAddr := 0, nValue := 16#BEEF);
rcoils(bExecute := st = 2, tTimeout := T#5s,
       sHost := '127.0.0.1', nTCPPort := 15089,
       nUnitID := 16#FF, nQuantity := 8, nMBAddr := 0,
       cbLength := 256);
rbad(bExecute := st = 3, tTimeout := T#5s,
     sHost := '127.0.0.1', nTCPPort := 15089,
     nUnitID := 16#FF, nQuantity := 2, nMBAddr := 99,
     cbLength := 256);
rwregs(bExecute := st = 4, tTimeout := T#5s,
       sHost := '127.0.0.1', nTCPPort := 15089,
       nUnitID := 16#FF, nReadQuantity := 2, nMBReadAddr := 0,
       nWriteQuantity := 1, nMBWriteAddr := 0,
       cbDestLength := 256, cbSrcLength := 2,
       pSrcData := wsrc);

IF st = 0 AND rregs.bDone THEN
    // func3 resp PDU data = bytecount + reg bytes
    IF rregs.bError = FALSE AND rregs.cbRead = 5 AND
       rregs.pData[0] = 4 AND rregs.pData[1] = 16#10 AND
       rregs.pData[2] = 16#00 AND rregs.pData[3] = 16#10 AND
       rregs.pData[4] = 16#01 THEN
        mask := mask + 1;
    END_IF;
    st := 1;
ELSIF st = 1 AND wsreg.bDone THEN
    IF wsreg.bError = FALSE AND wsreg.nErrId = 0 THEN
        mask := mask + 2;
    END_IF;
    st := 2;
ELSIF st = 2 AND rcoils.bDone THEN
    // func1 resp = bytecount(1) + 0xA5
    IF rcoils.bError = FALSE AND rcoils.cbRead = 2 AND
       rcoils.pData[0] = 1 AND rcoils.pData[1] = 16#A5 THEN
        mask := mask + 4;
    END_IF;
    st := 3;
ELSIF st = 3 AND rbad.bDone THEN
    // addr 99 -> server exception 2 -> nErrId = 16#8002
    IF rbad.bError = TRUE AND rbad.nErrId = 16#8002 THEN
        mask := mask + 8;
    END_IF;
    st := 4;
ELSIF st = 4 AND rwregs.bDone THEN
    IF rwregs.bError = FALSE AND rwregs.cbRead = 5 AND
       rwregs.pDestData[0] = 4 AND rwregs.pDestData[1] = 16#10 AND
       rwregs.pDestData[4] = 16#01 THEN
        mask := mask + 16;
    END_IF;
    st := 5;
END_IF;

scan_n := scan_n + 1;
END_PROGRAM

(* ---- tc2_motion_case.st ---- *)
PROGRAM Tc2MotionCase
VAR
    mask   AT %QD0 : DINT;
    st     : INT;
    ax     : FB_MotionAxis;
    axH    : UDINT;
    aStatus : DINT;
    aTgt   : DINT;
    aPos   : DINT;
    aVel   : DINT;
    sst    : DINT;
    gotEn  : BOOL;
END_VAR

// Deterministic simulated CiA402 axis exercised through the
// FB_MotionAxis builtin (tplc-motion service). One poll per scan
// advances dynamics; each state performs synchronous ops.
// DS402 object indices: 0x6040 cw, 0x6060 mode, 0x607A pos target,
// 0x60FF vel target. Controlword 0x001F = enable op + new setpoint.
ax.OP := 3;   // poll: advance all axes by the sim clock
ax();

IF st = 0 THEN
    // create: units/rev 1000, vmax 1000 u/s, accel/decel 5000 u/s^2
    ax.UNITS_PER_REV := 1000;
    ax.MAX_VEL := 1000;
    ax.MAX_ACCEL := 5000;
    ax.MAX_DECEL := 5000;
    ax.POS_MIN := -100000;
    ax.POS_MAX := 100000;
    ax.HOME_OFFSET := 0;
    ax.FOLLOW_WINDOW := 3;
    ax.FLAGS := 1;
    ax.OP := 1;
    ax();
    IF ax.AXIS <> 0 AND ax.STATUS = 0 THEN
        axH := ax.AXIS;
        mask := mask + 1;
    END_IF;
    st := 1;
ELSIF st = 1 THEN
    // mode = profile position (1)
    ax.OP := 5; ax.INDEX := 16#6060; ax.VALUE := 1; ax();
    IF ax.STATUS = 0 THEN mask := mask + 2; END_IF;
    st := 2;
ELSIF st = 2 THEN
    // target position = 500
    ax.OP := 5; ax.INDEX := 16#607A; ax.VALUE := 500; ax();
    IF ax.STATUS = 0 THEN mask := mask + 4; END_IF;
    st := 3;
ELSIF st = 3 THEN
    // controlword 0x001F: enable operation + new setpoint edge
    ax.OP := 5; ax.INDEX := 16#6040; ax.VALUE := 31; ax();
    IF ax.STATUS = 0 THEN mask := mask + 8; END_IF;
    st := 4;
ELSIF st = 4 THEN
    // wait for operation-enabled then the PP move to finish
    ax.OP := 6; ax.AXIS := axH; ax();
    aStatus := ax.STATUS;
    aTgt := ax.TARGET_REACHED;
    aPos := ax.POS_ACTUAL; aVel := ax.VEL_ACTUAL;
    sst := aStatus;
    IF sst = 39 AND NOT gotEn THEN
        gotEn := TRUE;
        mask := mask + 16;   // reached CiA402 OperationEnabled (0x27)
    END_IF;
    IF aTgt = 1 AND aPos >= 497 AND aPos <= 503 THEN
        mask := mask + 32;   // target reached within follow window
        st := 5;
    END_IF;
ELSIF st = 5 THEN
    // velocity mode: mode=2, target_vel=800 -> vel_actual ~800
    ax.OP := 5; ax.INDEX := 16#6060; ax.VALUE := 2; ax();
    ax.OP := 5; ax.INDEX := 16#60FF; ax.VALUE := 800; ax();
    st := 6;
ELSIF st = 6 THEN
    // wait for velocity to settle near 800 and position to move
    ax.OP := 6; ax.AXIS := axH; ax();
    aVel := ax.VEL_ACTUAL; aPos := ax.POS_ACTUAL;
    IF aVel >= 790 AND aVel <= 810 THEN
        mask := mask + 64;
        st := 7;
    END_IF;
ELSIF st = 7 THEN
    // error paths: bad object index read, bad mode write
    ax.OP := 4; ax.INDEX := 16#9999; ax();
    IF ax.STATUS < 0 THEN mask := mask + 128; END_IF;
    ax.OP := 5; ax.INDEX := 16#6060; ax.VALUE := 99; ax();
    IF ax.STATUS < 0 THEN mask := mask + 256; END_IF;
    // info on an invalid handle
    ax.OP := 6; ax.AXIS := 9999; ax();
    IF ax.STATUS < 0 THEN mask := mask + 512; END_IF;
    st := 8;
ELSIF st = 8 THEN
    // restore a valid mode, then destroy the axis
    ax.OP := 5; ax.INDEX := 16#6060; ax.VALUE := 1; ax.AXIS := axH; ax();
    ax.OP := 2; ax.AXIS := axH; ax();
    IF ax.STATUS = 0 THEN mask := mask + 1024; END_IF;
    st := 9;
ELSIF st = 9 THEN
    // info on the destroyed handle must fail
    ax.OP := 6; ax.AXIS := axH; ax();
    IF ax.STATUS < 0 THEN mask := mask + 2048; END_IF;
    st := 10;
END_IF;

END_PROGRAM

(* ---- tc2_mpbus_case.st ---- *)
// tc2_mpbus_case.st — wired MP-Bus e2e over a PTY slave fake
// (node 0x05).  Open, damper setpoint write -> ack, actual-pos
// read -> 0x80 (~50%), CMV read -> 0x42, close.
PROGRAM tc2_mpbus_case
VAR
    opn : FB_MpbusOpen;
    cls : FB_MpbusClose;
    dmp : MP_DamperLinearActuator;
    cmv : MP_CMV;
    st : INT;
    waitN : INT;
    mask AT %QD0 : UDINT;
    diag AT %QD4 : UDINT;
    hdl : UDINT;
END_VAR
    diag := st;
    IF st = 0 THEN
        mask := 0;
        opn.Execute := TRUE;
        opn.Path := '/tmp/mpb_pty';
        st := 1;
    ELSIF st = 1 THEN
        IF opn.Done THEN
            hdl := opn.PortHdl;
            opn.Execute := FALSE;
            mask := mask OR 1;        // bit0: serial open
            dmp.Execute := TRUE;
            dmp.PortHdl := hdl;
            dmp.DestAddr := 16#05;
            dmp.WriteSp := TRUE;
            dmp.Setpoint := 50.0;
            st := 2;
        END_IF;
        IF opn.Error THEN diag := 16#D0; st := 99; END_IF;
    ELSIF st = 2 THEN
        waitN := waitN + 1;
        IF dmp.Done THEN
            mask := mask OR 2;        // bit1: SP write ack
            st := 3;
        END_IF;
        IF dmp.Error THEN diag := 16#D1; st := 99; END_IF;
        IF waitN > 80 THEN diag := 16#D2; st := 99; END_IF;
    ELSIF st = 3 THEN
        // switch to actual-position read
        dmp.Execute := FALSE;
        waitN := 0;
        st := 4;
    ELSIF st = 4 THEN
        dmp.WriteSp := FALSE;
        dmp.Execute := TRUE;
        waitN := waitN + 1;
        IF dmp.Done THEN
            IF dmp.ActualPos > 45.0 AND dmp.ActualPos < 55.0 THEN
                mask := mask OR 4;    // bit2: actual pos ~50%
            END_IF;
            st := 5;
        END_IF;
        IF dmp.Error THEN diag := 16#D3; st := 99; END_IF;
        IF waitN > 80 THEN diag := 16#D4; st := 99; END_IF;
    ELSIF st = 5 THEN
        dmp.Execute := FALSE;
        cmv.Execute := TRUE;
        cmv.PortHdl := hdl;
        cmv.DestAddr := 16#05;
        cmv.Channel := 1;
        waitN := 0;
        st := 6;
    ELSIF st = 6 THEN
        waitN := waitN + 1;
        IF cmv.Done THEN
            IF cmv.Value = 16#42 THEN
                mask := mask OR 8;    // bit3: CMV value
            END_IF;
            cls.Execute := TRUE;
            cls.PortHdl := hdl;
            st := 7;
        END_IF;
        IF cmv.Error THEN diag := 16#D5; st := 99; END_IF;
        IF waitN > 80 THEN diag := 16#D6; st := 99; END_IF;
    ELSIF st = 7 THEN
        cmv.Execute := FALSE;
        IF cls.Done THEN
            mask := mask OR 16;       // bit4: close ok
            st := 8;
        END_IF;
        IF cls.Error THEN diag := 16#D7; st := 99; END_IF;
    END_IF;

    opn(); cls(); dmp(); cmv();
END_PROGRAM

(* ---- tc2_mqtt5_case.st ---- *)
// tc2_mqtt5_case.st — MQTT 5.0 client e2e over the python fake
// broker.  Connect via FB_IotMqtt5Client with connect properties,
// subscribe, publish, receive the echo, unsubscribe, disconnect.
PROGRAM tc2_mqtt5_case
VAR
    con : FB_IotMqtt5Client;
    dis : FB_IotMqttDisconnect;
    sub : FB_IotMqtt5Subscribe;
    unsub : FB_IotMqttUnsubscribe;
    pub : FB_IotMqttPublish;
    pub5 : FB_IotMqtt5Publish;
    rx  : FB_IotMqttReceive;
    rx5 : FB_IotMqtt5Receive;
    mq  : FB_IotMqtt5MessageQueue;
    up  : FB_IotMqtt5UserProperties;
    st : INT;
    waitN : INT;
    mask AT %QD0 : UDINT;
    hdl : UDINT;
END_VAR
    con(); dis(); sub(); unsub(); pub(); pub5(); rx(); rx5(); mq(); up();
    IF st = 0 THEN
        mask := 0;
        con.Execute := TRUE;
        con.HostName := '127.0.0.1';
        con.Port := 11883;
        con.CleanSession := TRUE;
        con.KeepAlive := 60;
        con.SessionExpiryS := 30;
        con.ReceiveMaximum := 10;
        con.TopicAliasMaximum := 4;
        con.RequestResponseInformation := TRUE;
        con.RequestProblemInformation := TRUE;
        st := 1;
    END_IF;

    IF st = 1 THEN
        IF con.Done THEN
            hdl := con.ConnectionHdl;
            con.Execute := FALSE;
            mask := mask + 1;         // bit0: v5 connected
            sub.Execute := TRUE;
            sub.ConnectionHdl := hdl;
            sub.TopicFilter := 'tplc/v5/#';
            sub.QoS := 0;
            sub.NoLocal := FALSE;
            sub.RetainAsPublished := FALSE;
            sub.RetainHandling := 0;
            sub.SubscriptionId := 7;
            sub.UserProperties := 'sk=sv';
            st := 2;
        END_IF;
        IF con.Error THEN mask := 16#DEAD; st := 99; END_IF;
    END_IF;

    IF st = 2 THEN
        IF sub.Done THEN
            sub.Execute := FALSE;
            mask := mask + 2;         // bit1: subscribed (v5 SUBACK)
            pub.Execute := TRUE;
            pub.ConnectionHdl := hdl;
            pub.Topic := 'tplc/v5/one';
            pub.Payload := 'm5';
            pub.QoS := 0;
            st := 3;
        END_IF;
        IF sub.Error THEN mask := 16#DEAD; st := 99; END_IF;
    END_IF;

    IF st = 3 THEN
        IF pub.Done THEN
            pub.Execute := FALSE;
            mask := mask + 4;         // bit2: published (v5 PUBLISH)
            waitN := 0;
            st := 4;
        END_IF;
        IF pub.Error THEN mask := 16#DEAD; st := 99; END_IF;
    END_IF;

    IF st = 4 THEN
        rx.Execute := TRUE;
        rx.ConnectionHdl := hdl;
        IF rx.Done AND rx.Message THEN
            rx.Execute := FALSE;
            IF rx.Topic = 'tplc/v5/one' AND rx.Payload = 'm5' THEN
                mask := mask + 8;     // bit3: echo received (v5)
                st := 50;
            END_IF;
        END_IF;
        IF rx.Error THEN mask := 16#DEAD; st := 99; END_IF;
        waitN := waitN + 1;
        IF waitN > 300 THEN mask := 16#DEAD; st := 99; END_IF;
    END_IF;

    IF st = 57 THEN
        IF pub5.Done THEN
            pub5.Execute := FALSE;
            waitN := 0;
            st := 58;
        END_IF;
        IF pub5.Error THEN mask := 16#DEAD; st := 99; END_IF;
    END_IF;

    IF st = 58 THEN
        IF mq.Queued > 0 THEN
            mq.DequeueReq := TRUE;
            st := 59;
        END_IF;
        waitN := waitN + 1;
        IF waitN > 300 THEN mask := 16#DEAD; st := 99; END_IF;
    END_IF;

    IF st = 59 THEN
        IF mq.HasMessage THEN
            mq.DequeueReq := FALSE;
            IF mq.Topic = 'tplc/v5/q/one'
               AND mq.Payload = 'qm'
               AND mq.MessageExpiryS = 10
               AND mq.ContentType = 'text/plain'
               AND mq.CorrelationData = 'qc'
               AND mq.CorrelationLen = 2
               AND mq.UserProperties = 'qk=qv' THEN
                mask := mask + 256;  // bit8: queued v5 props
                unsub.Execute := TRUE;
                unsub.ConnectionHdl := hdl;
                unsub.TopicFilter := 'tplc/v5/#';
                st := 5;
            ELSE
                mask := 16#DEAD; st := 99;
            END_IF;
        END_IF;
        waitN := waitN + 1;
        IF waitN > 300 THEN mask := 16#DEAD; st := 99; END_IF;
    END_IF;

    IF st = 5 THEN
        IF unsub.Done THEN
            unsub.Execute := FALSE;
            mask := mask + 16;        // bit4: unsubscribed
            dis.Execute := TRUE;
            dis.ConnectionHdl := hdl;
            st := 6;
        END_IF;
        IF unsub.Error THEN mask := 16#DEAD; st := 99; END_IF;
    END_IF;

    IF st = 50 THEN
        // stage user properties k1=v1 then k2=v2 via edge pulses;
        // ELSIF keeps one pulse per scan so up() sees each edge
        up.AddReq := TRUE;
        up.PropKey := 'k1';
        up.PropValue := 'v1';
        st := 51;
    ELSIF st = 51 THEN
        up.AddReq := FALSE;
        up.PropKey := 'k2';
        up.PropValue := 'v2';
        st := 52;
    ELSIF st = 52 THEN
        up.AddReq := TRUE;
        st := 53;
    ELSIF st = 53 THEN
        up.AddReq := FALSE;
        st := 54;
    END_IF;

    IF st = 54 THEN
        IF up.Count = 2 AND up.Encoded = 'k1=v1;k2=v2' THEN
            pub5.Execute := TRUE;
            pub5.ConnectionHdl := hdl;
            pub5.Topic := 'tplc/v5/props';
            pub5.Payload := 'withprops';
            pub5.QoS := 0;
            pub5.PayloadFormatUtf8 := TRUE;
            pub5.MessageExpiryS := 30;
            pub5.ContentType := 'application/json';
            pub5.ResponseTopic := 'tplc/v5/reply';
            pub5.CorrelationData := 'corr-1';
            pub5.UserProperties := up.Encoded;
            st := 55;
        ELSE
            mask := 16#F000 + up.Count * 16 + LEN(up.Encoded); st := 99;
        END_IF;
    END_IF;

    IF st = 55 THEN
        IF pub5.Done THEN
            pub5.Execute := FALSE;
            mask := mask + 64;        // bit6: v5 publish w/ props
            waitN := 0;
            st := 56;
        END_IF;
        IF pub5.Error THEN mask := 16#DEAD; st := 99; END_IF;
    END_IF;

    IF st = 56 THEN
        // pump the echo so the broker forwards the message; the
        // props themselves are verified broker-side via the log
        rx5.Execute := TRUE;
        rx5.ConnectionHdl := hdl;
        IF rx5.Done AND rx5.Message THEN
            rx5.Execute := FALSE;
            IF rx5.Topic = 'tplc/v5/props'
               AND rx5.PayloadFormatUtf8
               AND rx5.MessageExpiryS = 30
               AND rx5.ContentType = 'application/json'
               AND rx5.ResponseTopic = 'tplc/v5/reply'
               AND rx5.CorrelationData = 'corr-1'
               AND rx5.CorrelationLen = 6
               AND rx5.UserProperties = 'k1=v1;k2=v2' THEN
                mask := mask + 128; // bit7: props publish echoed
                // stage a queued v5 message with properties
                mq.Pump := TRUE;
                mq.ConnectionHdl := hdl;
                pub5.Execute := TRUE;
                pub5.Topic := 'tplc/v5/q/one';
                pub5.Payload := 'qm';
                pub5.PayloadFormatUtf8 := FALSE;
                pub5.MessageExpiryS := 10;
                pub5.ContentType := 'text/plain';
                pub5.ResponseTopic := '';
                pub5.CorrelationData := 'qc';
                pub5.UserProperties := 'qk=qv';
                st := 57;
            END_IF;
        END_IF;
        waitN := waitN + 1;
        IF waitN > 300 THEN mask := 16#DEAD; st := 99; END_IF;
    END_IF;

    IF st = 6 THEN
        IF dis.Done THEN
            mask := mask + 32;        // bit5: disconnected
            st := 7;
        END_IF;
        IF dis.Error THEN mask := 16#DEAD; st := 99; END_IF;
    END_IF;

    IF st = 7 THEN
        st := 8;
    END_IF;
END_PROGRAM

(* ---- tc2_mqtt5_req_case.st ---- *)
// tc2_mqtt5_req_case.st — MQTT5 request/response e2e: the fake
// broker runs in --responder mode and answers publishes on
// 'tplc/v5/req' that carry ResponseTopic + CorrelationData.
PROGRAM tc2_mqtt5_req_case
VAR
    con : FB_IotMqtt5Client;
    dis : FB_IotMqttDisconnect;
    req : FB_IotMqtt5RequestResponse;
    st : INT;
    waitN : INT;
    mask AT %QD0 : UDINT;
    hdl : UDINT;
END_VAR
    con(); dis(); req();
    IF st = 0 THEN
        mask := 0;
        con.Execute := TRUE;
        con.HostName := '127.0.0.1';
        con.Port := 11884;
        con.CleanSession := TRUE;
        con.KeepAlive := 60;
        st := 1;
    END_IF;

    IF st = 1 THEN
        IF con.Done THEN
            hdl := con.ConnectionHdl;
            con.Execute := FALSE;
            mask := mask + 1;         // bit0: v5 connected
            req.Execute := TRUE;
            req.ConnectionHdl := hdl;
            req.RequestTopic := 'tplc/v5/req';
            req.RequestPayload := 'ping';
            req.QoS := 0;
            req.ResponseTopic := 'tplc/v5/resp/in';
            req.CorrelationData := 'rc1';
            req.TimeoutScans := 400;
            st := 2;
        END_IF;
        IF con.Error THEN mask := 16#DEAD; st := 99; END_IF;
    END_IF;

    IF st = 2 THEN
        IF req.Done THEN
            req.Execute := FALSE;
            IF req.ResponsePayload = 'pong'
               AND req.ResponseTopicOut = 'tplc/v5/resp/in' THEN
                mask := mask + 2;     // bit1: correlated response
                dis.Execute := TRUE;
                dis.ConnectionHdl := hdl;
                st := 3;
            ELSE
                mask := 16#DEAD; st := 99;
            END_IF;
        END_IF;
        IF req.Error THEN mask := 16#DEAD; st := 99; END_IF;
        waitN := waitN + 1;
        IF waitN > 600 THEN mask := 16#DEAD; st := 99; END_IF;
    END_IF;

    IF st = 3 THEN
        IF dis.Done THEN
            mask := mask + 4;         // bit2: disconnected
            st := 4;
        END_IF;
        IF dis.Error THEN mask := 16#DEAD; st := 99; END_IF;
    END_IF;

    IF st = 4 THEN
        st := 5;
    END_IF;
END_PROGRAM

(* ---- tc2_mqtt_backoff_case.st ---- *)
// tc2_mqtt_backoff_case.st — exponential-backoff reconnect e2e.
// Connect + subscribe + echo, arm FB_IotMqttBackoff, then the io
// script kills the broker (connection drops), restarts it, and the
// host watchdog must reconnect with a doubling delay.  The case
// waits for the drop, waits for reconnect, resubscribes (subs are
// not restored), publishes a second message and receives its echo.
// mask bits 0..9 -> expect 0x3ff.
PROGRAM tc2_mqtt_backoff_case
VAR
    con  : FB_IotMqttClient;
    sub  : FB_IotMqttSubscribe;
    pub  : FB_IotMqttPublish;
    rx   : FB_IotMqttReceive;
    sts  : FB_IotMqttStatus;
    bo   : FB_IotMqttBackoff;
    sub2 : FB_IotMqttSubscribe;
    pub2 : FB_IotMqttPublish;
    rx2  : FB_IotMqttReceive;
    dis  : FB_IotMqttDisconnect;
    st : INT;
    waitN : INT;
    mask AT %QD0 : UDINT;
    hdl : UDINT;
END_VAR
    IF st = 0 THEN
        mask := 0;
        con.Execute := TRUE;
        con.HostName := '127.0.0.1';
        con.Port := 11885;
        con.CleanSession := TRUE;
        con.KeepAlive := 60;
        st := 1;
    END_IF;

    IF st = 1 THEN
        IF con.Done THEN
            hdl := con.ConnectionHdl;
            con.Execute := FALSE;
            mask := mask + 1;
            sub.Execute := TRUE;
            sub.ConnectionHdl := hdl;
            sub.TopicFilter := 'tplc/bo/#';
            sub.QoS := 0;
            st := 2;
        END_IF;
        IF con.Error THEN mask := 16#DEAD; st := 99; END_IF;
    END_IF;

    IF st = 2 THEN
        IF sub.Done THEN
            sub.Execute := FALSE;
            mask := mask + 2;
            pub.Execute := TRUE;
            pub.ConnectionHdl := hdl;
            pub.Topic := 'tplc/bo/a';
            pub.Payload := 'one';
            pub.QoS := 0;
            pub.RetainOn := FALSE;
            st := 3;
        END_IF;
        IF sub.Error THEN mask := 16#DEAD; st := 99; END_IF;
    END_IF;

    IF st = 3 THEN
        IF pub.Done THEN
            pub.Execute := FALSE;
            mask := mask + 4;
            // rx/sts start only after SUBACK+PUBLISH settled — a
            // concurrent MQTTClient_receive can steal the SUBACK
            // while subscribe waits for it
            rx.Execute := TRUE;
            rx.ConnectionHdl := hdl;
            sts.Execute := TRUE;
            sts.ConnectionHdl := hdl;
            waitN := 0;
            st := 4;
        END_IF;
        IF pub.Error THEN mask := 16#DEAD; st := 99; END_IF;
    END_IF;

    // first echo proves the baseline session works
    IF st = 4 THEN
        waitN := waitN + 1;
        IF rx.Message AND rx.Payload = 'one' THEN
            mask := mask + 8;
            bo.Execute := TRUE;
            bo.ConnectionHdl := hdl;
            bo.MinMs := 50;
            bo.MaxMs := 500;
            bo.Enable := TRUE;
            st := 5;
        END_IF;
        IF waitN > 600 THEN mask := 16#DEAD; st := 99; END_IF;
    END_IF;

    // arm the watchdog, then wait for the broker kill to surface
    IF st = 5 THEN
        IF bo.Done THEN
            bo.Execute := FALSE;
            mask := mask + 16;
            waitN := 0;
            st := 6;
        END_IF;
        IF bo.Error THEN mask := 16#DEAD; st := 99; END_IF;
    END_IF;

    // broker is dead: rx keeps polling so Paho observes the EOF
    IF st = 6 THEN
        waitN := waitN + 1;
        IF NOT sts.Connected THEN
            mask := mask + 32;
            waitN := 0;
            st := 7;
        END_IF;
        IF waitN > 800 THEN mask := 16#DEAD; st := 99; END_IF;
    END_IF;

    // broker restarted: watchdog reconnects (delay doubling)
    IF st = 7 THEN
        waitN := waitN + 1;
        IF sts.Connected THEN
            mask := mask + 64;
            sts.Execute := FALSE;
            rx.Execute := FALSE;
            sub2.Execute := TRUE;
            sub2.ConnectionHdl := hdl;
            sub2.TopicFilter := 'tplc/bo/#';
            sub2.QoS := 0;
            st := 8;
        END_IF;
        IF waitN > 1200 THEN mask := 16#DEAD; st := 99; END_IF;
    END_IF;

    IF st = 8 THEN
        IF sub2.Done THEN
            sub2.Execute := FALSE;
            mask := mask + 128;
            pub2.Execute := TRUE;
            pub2.ConnectionHdl := hdl;
            pub2.Topic := 'tplc/bo/b';
            pub2.Payload := 'two';
            pub2.QoS := 0;
            pub2.RetainOn := FALSE;
            rx2.Execute := TRUE;
            rx2.ConnectionHdl := hdl;
            waitN := 0;
            st := 9;
        END_IF;
        IF sub2.Error THEN mask := 16#DEAD; st := 99; END_IF;
    END_IF;

    IF st = 9 THEN
        waitN := waitN + 1;
        IF rx2.Message AND rx2.Payload = 'two' THEN
            mask := mask + 256;
            rx2.Execute := FALSE;
            dis.Execute := TRUE;
            dis.ConnectionHdl := hdl;
            st := 10;
        END_IF;
        IF waitN > 600 THEN mask := 16#DEAD; st := 99; END_IF;
    END_IF;

    IF st = 10 THEN
        IF dis.Done THEN
            mask := mask + 512;
            st := 11;
        END_IF;
        IF dis.Error THEN mask := 16#DEAD; st := 99; END_IF;
    END_IF;

    con(); sub(); pub(); rx(); sts(); bo();
    sub2(); pub2(); rx2(); dis();
END_PROGRAM

(* ---- tc2_mqtt_case.st ---- *)
// tc2_mqtt_case.st — MQTT client e2e over the python fake broker.
// Connect, publish retained, subscribe wildcard, receive the retained
// delivery (Retained=TRUE), publish live, receive the echo
// (Retained=FALSE), disconnect.  Then a second pair: a will-bearing
// client connects, a subscriber watches its will topic, the client
// aborts ungracefully (no DISCONNECT), and the broker's will delivery
// lands.  Also exercises F_MqttTopicMatch.
PROGRAM tc2_mqtt_case
VAR
    con : FB_IotMqttClient;
    dis : FB_IotMqttDisconnect;
    sub : FB_IotMqttSubscribe;
    pub : FB_IotMqttPublish;
    rx  : FB_IotMqttReceive;
    conW : FB_IotMqttClient;
    con2 : FB_IotMqttClient;
    sub2 : FB_IotMqttSubscribe;
    pub2 : FB_IotMqttPublish;
    rx2  : FB_IotMqttReceive;
    ab   : FB_IotMqttAbort;
    dis2 : FB_IotMqttDisconnect;
    st : INT;
    waitN : INT;
    mask AT %QD0 : UDINT;
    hdl : UDINT;
    hdlW : UDINT;
    hdl2 : UDINT;
END_VAR
    IF st = 0 THEN
        mask := 0;
        IF F_MqttTopicMatch('tplc/#', 'tplc/a/b')
           AND F_MqttTopicMatch('tplc/+/x', 'tplc/a/x')
           AND NOT F_MqttTopicMatch('tplc/+/x', 'tplc/a/y')
           AND F_MqttTopicMatch('a/b', 'a/b')
           AND NOT F_MqttTopicMatch('a/b', 'a/b/c') THEN
            mask := mask + 64;    // bit6: topic matcher
        END_IF;
        con.Execute := TRUE;
        con.HostName := '127.0.0.1';
        con.Port := 11883;
        con.CleanSession := TRUE;
        con.KeepAlive := 60;
        st := 1;
    END_IF;

    IF st = 1 THEN
        IF con.Done THEN
            hdl := con.ConnectionHdl;
            con.Execute := FALSE;
            mask := mask + 1;         // bit0: connected
            pub.Execute := TRUE;
            pub.ConnectionHdl := hdl;
            pub.Topic := 'tplc/keep';
            pub.Payload := 'saved';
            pub.QoS := 0;
            pub.RetainOn := TRUE;
            st := 2;
        END_IF;
        IF con.Error THEN mask := 16#DEAD; st := 99; END_IF;
    END_IF;

    IF st = 2 THEN
        IF pub.Done THEN
            mask := mask + 2;         // bit1: retained publish sent
            pub.Execute := FALSE;
            sub.Execute := TRUE;
            sub.ConnectionHdl := hdl;
            sub.TopicFilter := 'tplc/#';
            sub.QoS := 0;
            st := 3;
        END_IF;
        IF pub.Error THEN mask := 16#DEAD; st := 99; END_IF;
    END_IF;

    IF st = 3 THEN
        IF sub.Done THEN
            mask := mask + 4;         // bit2: subscribed
            sub.Execute := FALSE;
            rx.Execute := TRUE;
            rx.ConnectionHdl := hdl;
            st := 4;
        END_IF;
        IF sub.Error THEN mask := 16#DEAD; st := 99; END_IF;
    END_IF;

    // first message must be the broker's retained delivery
    IF st = 4 THEN
        waitN := waitN + 1;
        IF rx.Message THEN
            IF rx.Topic = 'tplc/keep' AND rx.Payload = 'saved'
               AND rx.Retained THEN
                mask := mask + 8;     // bit3: retained msg landed
            END_IF;
            // keep rx.Execute TRUE so st5 keeps polling for the echo
            pub.Execute := TRUE;
            pub.ConnectionHdl := hdl;
            pub.Topic := 'tplc/test';
            pub.Payload := 'hello';
            pub.QoS := 0;
            pub.RetainOn := FALSE;
            st := 5;
        END_IF;
        IF rx.Error THEN mask := 16#DEAD; st := 99; END_IF;
        IF waitN > 400 THEN
            rx.Execute := FALSE;
            dis.Execute := TRUE;
            dis.ConnectionHdl := hdl;
            st := 6;
        END_IF;
    END_IF;

    // second message is the live echo of our publish
    IF st = 5 THEN
        waitN := waitN + 1;
        IF rx.Message THEN
            IF rx.Topic = 'tplc/test' AND rx.Payload = 'hello'
               AND NOT rx.Retained THEN
                mask := mask + 16;    // bit4: live echo, not retained
                rx.Execute := FALSE;
                dis.Execute := TRUE;
                dis.ConnectionHdl := hdl;
                st := 6;
            END_IF;
            // non-matching messages (e.g. a repeated retained
            // delivery) are consumed and polling continues
        END_IF;
        IF rx.Error THEN mask := 16#DEAD; st := 99; END_IF;
        IF waitN > 400 THEN
            rx.Execute := FALSE;
            dis.Execute := TRUE;
            dis.ConnectionHdl := hdl;
            st := 6;
        END_IF;
    END_IF;

    IF st = 6 THEN
        IF dis.Done THEN
            mask := mask + 32;        // bit5: disconnected
            conW.Execute := TRUE;
            conW.HostName := '127.0.0.1';
            conW.Port := 11883;
            conW.CleanSession := TRUE;
            conW.KeepAlive := 60;
            conW.WillTopic := 'tplc/will';
            conW.WillPayload := 'gone';
            conW.WillQoS := 0;
            conW.WillRetain := FALSE;
            st := 7;
        END_IF;
        IF dis.Error THEN mask := 16#DEAD; st := 99; END_IF;
    END_IF;

    // will client connected -> bring up the watcher connection
    IF st = 7 THEN
        IF conW.Done THEN
            hdlW := conW.ConnectionHdl;
            conW.Execute := FALSE;
            mask := mask + 128;       // bit7: will client connected
            con2.Execute := TRUE;
            con2.HostName := '127.0.0.1';
            con2.Port := 11883;
            con2.CleanSession := TRUE;
            con2.KeepAlive := 60;
            st := 8;
        END_IF;
        IF conW.Error THEN mask := 16#DEAD; st := 99; END_IF;
    END_IF;

    IF st = 8 THEN
        IF con2.Done THEN
            hdl2 := con2.ConnectionHdl;
            con2.Execute := FALSE;
            sub2.Execute := TRUE;
            sub2.ConnectionHdl := hdl2;
            sub2.TopicFilter := 'tplc/will';
            sub2.QoS := 0;
            st := 9;
        END_IF;
        IF con2.Error THEN mask := 16#DEAD; st := 99; END_IF;
    END_IF;

    IF st = 9 THEN
        IF sub2.Done THEN
            sub2.Execute := FALSE;
            mask := mask + 256;       // bit8: will topic subscribed
            // sanity: conn2 rx path works before the abort — publish
            // a ping to its own subscription (echo arrives as 'ping',
            // ignored by the will check in st11)
            pub2.Execute := TRUE;
            pub2.ConnectionHdl := hdl2;
            pub2.Topic := 'tplc/will';
            pub2.Payload := 'ping';
            pub2.QoS := 0;
            pub2.RetainOn := FALSE;
            rx2.Execute := TRUE;
            rx2.ConnectionHdl := hdl2;
            waitN := 0;
            st := 10;
        END_IF;
        IF sub2.Error THEN mask := 16#DEAD; st := 99; END_IF;
    END_IF;

    // wait for the self-ping echo, then abort the will client
    IF st = 10 THEN
        waitN := waitN + 1;
        IF rx2.Message AND rx2.Payload = 'ping' THEN
            mask := mask + 512;       // bit9: conn2 rx path verified
            ab.Execute := TRUE;
            ab.ConnectionHdl := hdlW;
            st := 13;
        END_IF;
        IF rx2.Error THEN mask := 16#DEAD; st := 99; END_IF;
        IF pub2.Error THEN mask := 16#DEAD; st := 99; END_IF;
        IF waitN > 400 THEN mask := 16#DEAD; st := 99; END_IF;
    END_IF;

    // ungraceful drop: no DISCONNECT, broker must fire the will
    IF st = 13 THEN
        IF ab.Done THEN
            ab.Execute := FALSE;
            waitN := 0;
            st := 11;
        END_IF;
        IF ab.Error THEN mask := 16#DEAD; st := 99; END_IF;
    END_IF;

    IF st = 11 THEN
        waitN := waitN + 1;
        IF rx2.Message THEN
            IF rx2.Topic = 'tplc/will' AND rx2.Payload = 'gone' THEN
                mask := mask + 1024;  // bit10: will delivered
                rx2.Execute := FALSE;
                dis2.Execute := TRUE;
                dis2.ConnectionHdl := hdl2;
                st := 12;
            END_IF;
        END_IF;
        IF rx2.Error THEN mask := 16#DEAD; st := 99; END_IF;
        IF waitN > 400 THEN mask := 16#DEAD; st := 99; END_IF;
    END_IF;

    IF st = 12 THEN
        IF dis2.Done THEN
            mask := mask + 2048;      // bit11: watcher disconnected
            st := 14;
        END_IF;
        IF dis2.Error THEN mask := 16#DEAD; st := 99; END_IF;
    END_IF;

    con(); dis(); sub(); pub(); rx();
    conW(); con2(); sub2(); pub2(); rx2(); ab(); dis2();
END_PROGRAM

(* ---- tc2_mqtt_queue_case.st ---- *)
// tc2_mqtt_queue_case.st — MQTT message-queue e2e over the python
// fake broker: connect, subscribe tplc/q/#, pump three published
// messages into FB_IotMqttMessageQueue, dequeue them FIFO, reset the
// queue, publish+dequeue a fourth, disconnect.
// NOTE: separate FB_IotMqttPublish instances per message — the FBs
// are edge-triggered and same-scan re-arming never produces an edge.
PROGRAM tc2_mqtt_queue_case
VAR
    con : FB_IotMqttClient;
    dis : FB_IotMqttDisconnect;
    sub : FB_IotMqttSubscribe;
    pub1 : FB_IotMqttPublish;
    pub2 : FB_IotMqttPublish;
    pub3 : FB_IotMqttPublish;
    pub4 : FB_IotMqttPublish;
    sub2 : FB_IotMqttSubscribe;
    pub5 : FB_IotMqttPublish;
    q : FB_IotMqttMessageQueue;
    st : INT;
    waitN : INT;
    dqPend : INT;
    dqN : INT;
    mask AT %QD0 : UDINT;
    hdl : UDINT;
END_VAR
    IF st = 0 THEN
        mask := 0;
        waitN := 0;
        con.Execute := TRUE;
        con.HostName := '127.0.0.1';
        con.Port := 11883;
        con.CleanSession := TRUE;
        con.KeepAlive := 60;
        st := 1;
    END_IF;

    IF st = 1 THEN
        IF con.Done THEN
            hdl := con.ConnectionHdl;
            con.Execute := FALSE;
            mask := mask + 1;              // bit0: connected
            sub.Execute := TRUE;
            sub.ConnectionHdl := hdl;
            sub.TopicFilter := 'tplc/q/#';
            sub.QoS := 0;
            q.Pump := TRUE;
            q.ConnectionHdl := hdl;
            st := 2;
        END_IF;
        IF con.Error THEN mask := 16#DEAD; st := 99; END_IF;
    END_IF;

    IF st = 2 THEN
        IF sub.Done THEN
            sub.Execute := FALSE;
            mask := mask + 2;              // bit1: subscribed
            pub1.Execute := TRUE;
            pub1.ConnectionHdl := hdl;
            pub1.Topic := 'tplc/q/one';
            pub1.Payload := 'm1';
            pub1.QoS := 0;
            st := 3;
        END_IF;
        IF sub.Error THEN mask := 16#DEAD; st := 99; END_IF;
    END_IF;

    IF st = 3 THEN
        IF pub1.Done THEN
            pub1.Execute := FALSE;
            pub2.Execute := TRUE;
            pub2.ConnectionHdl := hdl;
            pub2.Topic := 'tplc/q/two';
            pub2.Payload := 'm2';
            pub2.QoS := 0;
            st := 4;
        END_IF;
        IF pub1.Error THEN mask := 16#DEAD; st := 99; END_IF;
    END_IF;

    IF st = 4 THEN
        IF pub2.Done THEN
            pub2.Execute := FALSE;
            pub3.Execute := TRUE;
            pub3.ConnectionHdl := hdl;
            pub3.Topic := 'tplc/q/three';
            pub3.Payload := 'm3';
            pub3.QoS := 0;
            st := 5;
        END_IF;
        IF pub2.Error THEN mask := 16#DEAD; st := 99; END_IF;
    END_IF;

    IF st = 5 THEN
        IF pub3.Done THEN
            pub3.Execute := FALSE;
            waitN := 0;
            st := 6;
        END_IF;
        IF pub3.Error THEN mask := 16#DEAD; st := 99; END_IF;
    END_IF;

    // wait for the pump to collect all three messages
    IF st = 6 THEN
        waitN := waitN + 1;
        IF q.Queued >= 3 THEN
            mask := mask + 4;              // bit2: queue filled
            dqN := 0;
            dqPend := 0;
            st := 7;
        ELSIF waitN > 300 THEN
            mask := 16#DEAD; st := 99;
        END_IF;
        IF q.Error THEN mask := 16#DEAD; st := 99; END_IF;
    END_IF;

    // dequeue x3 with a one-scan request pulse; outputs are checked
    // the scan after each request
    IF st = 7 THEN
        IF dqPend = 0 THEN
            q.DequeueReq := TRUE;
            dqPend := 1;
        ELSE
            q.DequeueReq := FALSE;
            IF q.HasMessage THEN
                dqN := dqN + 1;
                IF dqN = 1 AND q.Topic = 'tplc/q/one'
                   AND q.Payload = 'm1' THEN
                    mask := mask + 8;       // bit3: FIFO m1
                END_IF;
                IF dqN = 2 AND q.Topic = 'tplc/q/two'
                   AND q.Payload = 'm2' THEN
                    mask := mask + 16;      // bit4: FIFO m2
                END_IF;
                IF dqN = 3 AND q.Topic = 'tplc/q/three'
                   AND q.Payload = 'm3' THEN
                    mask := mask + 32;      // bit5: FIFO m3
                END_IF;
            END_IF;
            dqPend := 0;
            IF dqN >= 3 THEN st := 8; END_IF;
        END_IF;
        IF q.Error THEN mask := 16#DEAD; st := 99; END_IF;
    END_IF;

    // queue must now be empty; reset and verify
    IF st = 8 THEN
        IF q.Queued = 0 THEN
            mask := mask + 64;             // bit6: drained
            q.ResetReq := TRUE;
            st := 9;
        ELSE
            waitN := waitN + 1;
            IF waitN > 300 THEN mask := 16#DEAD; st := 99; END_IF;
        END_IF;
    END_IF;

    IF st = 9 THEN
        q.ResetReq := FALSE;
        pub4.Execute := TRUE;
        pub4.ConnectionHdl := hdl;
        pub4.Topic := 'tplc/q/four';
        pub4.Payload := 'm4';
        pub4.QoS := 0;
        waitN := 0;
        st := 10;
    END_IF;

    // pump refills; wait for the fourth message then dequeue it
    IF st = 10 THEN
        waitN := waitN + 1;
        IF q.Queued >= 1 THEN
            dqPend := 0;
            st := 11;
        ELSIF waitN > 300 THEN
            mask := 16#DEAD; st := 99;
        END_IF;
    END_IF;

    IF st = 11 THEN
        IF dqPend = 0 THEN
            q.DequeueReq := TRUE;
            dqPend := 1;
        ELSE
            q.DequeueReq := FALSE;
            IF q.HasMessage AND q.Topic = 'tplc/q/four'
               AND q.Payload = 'm4' THEN
                mask := mask + 128;       // bit7: post-reset msg
            END_IF;
            dqPend := 0;
            st := 12;
        END_IF;
    END_IF;

    // QoS2 stage: subscribe at granted qos2, publish qos2, the
    // PUBREC/PUBREL/PUBCOMP handshake runs inside Paho + the fake
    // broker; the dequeued message must report QoS=2
    IF st = 12 THEN
        sub2.Execute := TRUE;
        sub2.ConnectionHdl := hdl;
        sub2.TopicFilter := 'tplc/q2/#';
        sub2.QoS := 2;
        st := 14;
    END_IF;

    IF st = 14 THEN
        IF sub2.Done THEN
            sub2.Execute := FALSE;
            pub5.Execute := TRUE;
            pub5.ConnectionHdl := hdl;
            pub5.Topic := 'tplc/q2/five';
            pub5.Payload := 'm5';
            pub5.QoS := 2;
            waitN := 0;
            st := 15;
        END_IF;
        IF sub2.Error THEN mask := 16#DEAD; st := 99; END_IF;
    END_IF;

    IF st = 15 THEN
        IF pub5.Done THEN
            pub5.Execute := FALSE;
            waitN := 0;
            st := 16;
        END_IF;
        IF pub5.Error THEN mask := 16#DEAD; st := 99; END_IF;
    END_IF;

    IF st = 16 THEN
        waitN := waitN + 1;
        IF q.Queued >= 1 THEN
            dqPend := 0;
            st := 17;
        ELSIF waitN > 300 THEN
            mask := 16#DEAD; st := 99;
        END_IF;
    END_IF;

    IF st = 17 THEN
        IF dqPend = 0 THEN
            q.DequeueReq := TRUE;
            dqPend := 1;
        ELSE
            q.DequeueReq := FALSE;
            IF q.HasMessage AND q.Topic = 'tplc/q2/five'
               AND q.Payload = 'm5' AND q.QoS = 2 THEN
                mask := mask + 512;       // bit9: qos2 delivery
            END_IF;
            dqPend := 0;
            st := 18;
        END_IF;
    END_IF;

    IF st = 18 THEN
        dis.Execute := TRUE;
        dis.ConnectionHdl := hdl;
        st := 19;
    END_IF;

    IF st = 19 THEN
        IF dis.Done THEN
            dis.Execute := FALSE;
            mask := mask + 1024;           // bit10: disconnected
            st := 99;
        END_IF;
        IF dis.Error THEN mask := 16#DEAD; st := 99; END_IF;
    END_IF;

    con(); dis(); sub(); pub1(); pub2(); pub3(); pub4(); sub2(); pub5(); q();
END_PROGRAM

(* ---- tc2_mqtt_tls_case.st ---- *)
// tc2_mqtt_tls_case.st — MQTT over TLS e2e against the python fake
// broker's --tls mode.  conn1 uses UseTls+TlsInsecure (skip verify,
// self-signed broker); conn2 verifies against TlsCaFile (the
// broker's self-signed cert doubles as its own CA).  Each
// connection: CONNECT -> SUBSCRIBE -> PUBLISH -> receive echo ->
// DISCONNECT; conn1 also polls FB_IotMqttStatus for the
// broker-message age.  mask bits 0..10 -> expect 0x7ff.
PROGRAM tc2_mqtt_tls_case
VAR
    con1 : FB_IotMqttClient;
    sub1 : FB_IotMqttSubscribe;
    pub1 : FB_IotMqttPublish;
    rx1  : FB_IotMqttReceive;
    dis1 : FB_IotMqttDisconnect;
    con2 : FB_IotMqttClient;
    sub2 : FB_IotMqttSubscribe;
    pub2 : FB_IotMqttPublish;
    rx2  : FB_IotMqttReceive;
    dis2 : FB_IotMqttDisconnect;
    sts  : FB_IotMqttStatus;
    st : INT;
    waitN : INT;
    mask AT %QD0 : UDINT;
    hdl1 : UDINT;
    hdl2 : UDINT;
END_VAR
    IF st = 0 THEN
        mask := 0;
        con1.Execute := TRUE;
        con1.HostName := '127.0.0.1';
        con1.Port := 11884;
        con1.CleanSession := TRUE;
        con1.KeepAlive := 60;
        con1.UseTls := TRUE;
        con1.TlsInsecure := TRUE;
        st := 1;
    END_IF;

    IF st = 1 THEN
        IF con1.Done THEN
            hdl1 := con1.ConnectionHdl;
            con1.Execute := FALSE;
            mask := mask + 1;
            sub1.Execute := TRUE;
            sub1.ConnectionHdl := hdl1;
            sub1.TopicFilter := 'tplc/tls/#';
            sub1.QoS := 0;
            st := 2;
        END_IF;
        IF con1.Error THEN mask := 16#DEAD; st := 99; END_IF;
    END_IF;

    IF st = 2 THEN
        IF sub1.Done THEN
            sub1.Execute := FALSE;
            mask := mask + 2;
            pub1.Execute := TRUE;
            pub1.ConnectionHdl := hdl1;
            pub1.Topic := 'tplc/tls/a';
            pub1.Payload := 'secure1';
            pub1.QoS := 0;
            pub1.RetainOn := FALSE;
            st := 3;
        END_IF;
        IF sub1.Error THEN mask := 16#DEAD; st := 99; END_IF;
    END_IF;

    IF st = 3 THEN
        IF pub1.Done THEN
            pub1.Execute := FALSE;
            mask := mask + 4;
            rx1.Execute := TRUE;
            rx1.ConnectionHdl := hdl1;
            waitN := 0;
            st := 4;
        END_IF;
        IF pub1.Error THEN mask := 16#DEAD; st := 99; END_IF;
    END_IF;

    IF st = 4 THEN
        waitN := waitN + 1;
        IF rx1.Message THEN
            IF rx1.Topic = 'tplc/tls/a' AND rx1.Payload = 'secure1' THEN
                mask := mask + 8;
                rx1.Execute := FALSE;
                sts.Execute := TRUE;
                sts.ConnectionHdl := hdl1;
                st := 12;
            END_IF;
        END_IF;
        IF rx1.Error THEN mask := 16#DEAD; st := 99; END_IF;
        IF waitN > 400 THEN mask := 16#DEAD; st := 99; END_IF;
    END_IF;

    // status poll right after the echo: connected and the
    // broker-message age is fresh (the echo just landed)
    IF st = 12 THEN
        IF sts.Connected
           AND sts.TimeSinceLastBrokerMsgMs < 60000 THEN
            mask := mask + 1024;
            sts.Execute := FALSE;
            dis1.Execute := TRUE;
            dis1.ConnectionHdl := hdl1;
            st := 5;
        END_IF;
        IF sts.Error THEN mask := 16#DEAD; st := 99; END_IF;
    END_IF;

    IF st = 5 THEN
        IF dis1.Done THEN
            dis1.Execute := FALSE;
            mask := mask + 16;
            con2.Execute := TRUE;
            con2.HostName := '127.0.0.1';
            con2.Port := 11884;
            con2.CleanSession := TRUE;
            con2.KeepAlive := 60;
            con2.UseTls := TRUE;
            con2.TlsInsecure := FALSE;
            con2.TlsCaFile := '/tmp/tplc_mqtt_tls/cert.pem';
            st := 6;
        END_IF;
        IF dis1.Error THEN mask := 16#DEAD; st := 99; END_IF;
    END_IF;

    IF st = 6 THEN
        IF con2.Done THEN
            hdl2 := con2.ConnectionHdl;
            con2.Execute := FALSE;
            mask := mask + 32;
            sub2.Execute := TRUE;
            sub2.ConnectionHdl := hdl2;
            sub2.TopicFilter := 'tplc/tls/#';
            sub2.QoS := 0;
            st := 7;
        END_IF;
        IF con2.Error THEN mask := 16#DEAD; st := 99; END_IF;
    END_IF;

    IF st = 7 THEN
        IF sub2.Done THEN
            sub2.Execute := FALSE;
            mask := mask + 64;
            pub2.Execute := TRUE;
            pub2.ConnectionHdl := hdl2;
            pub2.Topic := 'tplc/tls/b';
            pub2.Payload := 'secure2';
            pub2.QoS := 0;
            pub2.RetainOn := FALSE;
            st := 8;
        END_IF;
        IF sub2.Error THEN mask := 16#DEAD; st := 99; END_IF;
    END_IF;

    IF st = 8 THEN
        IF pub2.Done THEN
            pub2.Execute := FALSE;
            mask := mask + 128;
            rx2.Execute := TRUE;
            rx2.ConnectionHdl := hdl2;
            waitN := 0;
            st := 9;
        END_IF;
        IF pub2.Error THEN mask := 16#DEAD; st := 99; END_IF;
    END_IF;

    IF st = 9 THEN
        waitN := waitN + 1;
        IF rx2.Message THEN
            IF rx2.Topic = 'tplc/tls/b' AND rx2.Payload = 'secure2' THEN
                mask := mask + 256;
                rx2.Execute := FALSE;
                dis2.Execute := TRUE;
                dis2.ConnectionHdl := hdl2;
                st := 10;
            END_IF;
        END_IF;
        IF rx2.Error THEN mask := 16#DEAD; st := 99; END_IF;
        IF waitN > 400 THEN mask := 16#DEAD; st := 99; END_IF;
    END_IF;

    IF st = 10 THEN
        IF dis2.Done THEN
            mask := mask + 512;
            st := 11;
        END_IF;
        IF dis2.Error THEN mask := 16#DEAD; st := 99; END_IF;
    END_IF;

    con1(); sub1(); pub1(); rx1(); dis1(); sts();
    con2(); sub2(); pub2(); rx2(); dis2();
END_PROGRAM
